(* IEC 61131-3 sources: ConveyorControl-with-PLC/4E_Gruppe1_Graf_Projekt1/Class/SafetyManager (part 3) *)

                    // change the command, because now we forward it to the receiver
                    pPara^.uiCmd := CMD_SM_SDO_TO_MODULE;

                    pHelpSafety^.pThis^.NewInst(pPara, #MyResult);
                    return;
                  else
                    pHelpSafety := pHelpSafety^.pNext;
                  end_if;
                end_while;
              end_if;
            end_if;

            pHelpPdo := pHelpPdo^.pNext;
          end_while;

          pHelpConfig := pHelpConfig^.pNext;
        end_while;
      end_if;
    end_if;

    // check if there is any interface frame domain optional and not available
    pHelpManaging := pFirstManagingInterfaceComponent;
    while pHelpManaging do
      if (pHelpManaging^.InfoBits.IsSynchron = 0) & (pHelpManaging^.InfoBits.IsOptional = 1) then
        // found one => no error here
        return;
      end_if;

      pHelpManaging := pHelpManaging^.pNext;
    end_while;

    // no optional interface domains missing => must be an error
    LogError("(SafetyManager::CheckTopSDO) Couldn't find InterfaceCRC. Check SafetyDesigner projects, maybe the interface variables do not match.");
    LogValue(pString:="SrcAddr: {0} / InterfaceCRC: {1}", Value:=pDO^.SrcAdr, Value2:=InterfaceCRC);
    ClassState := -8;

  // check if it's a local interface frame and we have no interface frame domains
  elsif (pCompDestPath^ = INTERFACE_CRC_MODE) then
    // after the mode byte we find the interface CRC
    InterfaceCRC := ((pCompDestPath + 1)$^HDINT)^;

    // search for the CRC
    pHelpSafety := NIL;
    if LocalIFNo then
      for i := 0 to (LocalIFNo-1) do
        if aLocalIFs[i].InterfaceCRC = InterfaceCRC then
          // found it
          pHelpSafety := aLocalIFs[i].pSafetyModule;
          exit;
        end_if;
      end_for;
    end_if;

    if pHelpSafety then
      // change the command, because now we forward it to the receiver
      pPara^.uiCmd := CMD_SM_SDO_TO_MODULE;

      pHelpSafety^.pThis^.NewInst(pPara, #MyResult);
    else
      // check the slave modules if there is one with the interface frame we need
      TargetSafetyNbr := 0;
      pHelpConfig := pConfigs;
      while pHelpConfig do
        pHelpSlave := pHelpConfig^.pFirstSlaveCfg;
        while pHelpSlave do

          if (pHelpSlave^.SlaveInfo.Info.IsInterface) & (pHelpSlave^.SlaveInfo.InterfaceCRC = InterfaceCRC) then
            // we have to add some additional information to the message

            (*
              Memory structure:
                1 Byte destination domain
                1 Byte IsInterfaceFrame (0/1)
                2 Byte length of uncompressed path
                x Byte uncompressed path
                x Byte SDO message
            *)

            MyPara.uiCmd := CMD_SM_TOP_SDO_TO_MODULE;
            MyPara.aPara[0] := sizeof(USINT) + sizeof(BOOL) + sizeof(UINT) + pHelpSlave^.SlaveInfo.PathLen + pPara^.aPara[0];

            if ud_SizeTempMemCy >= MyPara.aPara[0]$UDINT then
              pTempMem := pTempMemCy$^USINT;
            else
              LogError("(SafetyManager::CheckTopSDO) Temporary memory for cyclic task is too small!");
              LogValue(pString:="AvaliableMem: {0} / NeededMem: {1}", Value:=ud_SizeTempMemCy, Value2:=MyPara.aPara[0]$UDINT);
              return;
            end_if;

            TmpPathLen := pHelpSlave^.SlaveInfo.PathLen; // save some time with this local variable
            DomainChangeFound := FALSE;
            pHelp := pHelpSlave^.SlaveInfo.pPath + TmpPathLen - 2; // pointer on penultimate byte of path
            // search from the end for the last domain change
            for i := (TmpPathLen-2) to 3 by -1 do
              if pHelp^ = HWT_ESCAPE_DOMAIN then
                DomainChangeFound := TRUE;
                DestDomain := (pHelp + 1)^;
                exit;
              end_if;

              pHelp -= sizeof(USINT);
            end_for;

            // if there was no domainchange
            if DomainChangeFound = FALSE then
              // the master is the Dest
              DestDomain := (pHelpSlave^.SlaveInfo.pPath + 2)^;
            end_if;

            pHelp := pTempMem;

            // destination domain
            pHelp^ := DestDomain;
            pHelp += sizeof(USINT);

            // is it for an interface frame?
            pHelp^$BOOL := TRUE;
            pHelp += sizeof(BOOL);

            // length of uncompressed path
            pHelp^$UINT := TmpPathLen;
            pHelp += sizeof(UINT);

            // uncompressed path
            _memcpy(ptr1:=pHelp, ptr2:=pHelpSlave^.SlaveInfo.pPath, cntr:=TmpPathLen);
            pHelp += TmpPathLen;

            // SDO message
            _memcpy(ptr1:=pHelp, ptr2:=pDO, cntr:=pPara^.aPara[0]$UDINT);

            MyPara.aPara[1] := pTempMem$DINT;

            NewInst(#MyPara, #MyResult);

            // path can exist only once in a system
            return;
          end_if;

          pHelpSlave := pHelpSlave^.pNext;
        end_while;

        pHelpModule := pHelpConfig^.pFirstModuleCfg;
        while pHelpModule do
          if pHelpModule^.ModuleInfo.InterfaceCRC = InterfaceCRC then
            // if we found our target => forward the SDO to it
            TargetSafetyNbr := pHelpModule^.ModuleInfo.SafetyNbr;

            pHelpSafety := pFirstSafetyComponent;
            while pHelpSafety do
              // we compare the safety number
              if pHelpSafety^.SafetyNbr = TargetSafetyNbr then
                // change the command, because now we forward it to the receiver
                pPara^.uiCmd := CMD_SM_SDO_TO_MODULE;

                pHelpSafety^.pThis^.NewInst(pPara, #MyResult);

                return;
              end_if;

              pHelpSafety := pHelpSafety^.pNext;
            end_while;
          end_if;

          pHelpModule := pHelpModule^.pNext;
        end_while;

        pHelpConfig := pHelpConfig^.pNext;
      end_while;

      LogError("(SafetyManager::CheckTopSDO) Couldn't find target of SDO via TOP (Local Interface Frame)");
      LogValue(pString:="SrcAddr: {0} / InterfaceCRC: {1}", Value:=pDO^.SrcAdr, Value2:=InterfaceCRC);
    end_if;
  else
    // check if we have a module with this path
    pHelpConfig := pConfigs;
    while pHelpConfig do
      pHelpModule := pHelpConfig^.pFirstModuleCfg;
      while pHelpModule do
        if (To_StdLib.MemCmp(pCompDestPath, pHelpModule^.ModuleInfo.pCompPath, pHelpModule^.ModuleInfo.CompPathLen) = 0) then
          // we have to add some additional information to the message

          (*
            Memory structure:
              1 Byte destination domain
              1 Byte IsInterfaceFrame (0/1)
              2 Byte length of uncompressed path
              x Byte uncompressed path
              x Byte SDO message
          *)

          TmpPathLen := pHelpModule^.ModuleInfo.PathLen; // save some time with this local variable
          MyPara.uiCmd := CMD_SM_TOP_SDO_TO_MODULE;
          MyPara.aPara[0] := sizeof(USINT) + sizeof(BOOL) + sizeof(UINT) + TmpPathLen + pPara^.aPara[0];
          if ud_SizeTempMemCy >= MyPara.aPara[0]$UDINT then
            pTempMem := pTempMemCy$^USINT;
          else
            LogError("(SafetyManager::CheckTopSDO) Temporary memory for cyclic task is too small!");
            LogValue(pString:="AvaliableMem: {0} / NeededMem: {1}", Value:=ud_SizeTempMemCy, Value2:=MyPara.aPara[0]$UDINT);
            return;
          end_if;

          DomainChangeFound := FALSE;
          pHelp := pHelpModule^.ModuleInfo.pPath + TmpPathLen - 2; // pointer on penultimate byte of path
          // search from the end for the last domain change
          for i := (TmpPathLen-2) to 3 by -1 do
            if pHelp^ = HWT_ESCAPE_DOMAIN then
              DomainChangeFound := TRUE;
              DestDomain := (pHelp + 1)^;
              exit;
            end_if;

            pHelp -= sizeof(USINT);
          end_for;

          // if there was no domainchange
          if DomainChangeFound = FALSE then
            // the master is the Dest
            DestDomain := (pHelpModule^.ModuleInfo.pPath + 2)^;
          end_if;

          pHelp := pTempMem;

          // destination domain
          pHelp^ := DestDomain;
          pHelp += sizeof(USINT);

          // is it for an interface frame?
          pHelp^$BOOL := FALSE;
          pHelp += sizeof(BOOL);

          // length of uncompressed path
          pHelp^$UINT := TmpPathLen;
          pHelp += sizeof(UINT);

          // uncompressed path
          _memcpy(ptr1:=pHelp, ptr2:=pHelpModule^.ModuleInfo.pPath, cntr:=TmpPathLen);
          pHelp += TmpPathLen;

          // SDO message
          _memcpy(ptr1:=pHelp, ptr2:=pDO, cntr:=pPara^.aPara[0]$UDINT);

          MyPara.aPara[1] := pTempMem$DINT;

          NewInst(#MyPara, #MyResult);

          // path can exist only once in a system
          return;
        end_if;

        pHelpModule := pHelpModule^.pNext;
      end_while;

      if pHelpConfig^.SafetyNbr = pDO^.SrcAdr then
        pHelpSlave := pHelpConfig^.pFirstSlaveCfg;
        while pHelpSlave do
          if (To_StdLib.MemCmp(pCompDestPath, pHelpSlave^.SlaveInfo.pCompPath, pHelpSlave^.SlaveInfo.CompPathLen) = 0) then
            // we have to add some additional information to the message

            (*
              Memory structure:
                1 Byte destination domain
                1 Byte IsInterfaceFrame (0/1)
                2 Byte length of uncompressed path
                x Byte uncompressed path
                x Byte SDO message
            *)

            TmpPathLen := pHelpSlave^.SlaveInfo.PathLen; // save some time with this local variable
            MyPara.uiCmd := CMD_SM_TOP_SDO_TO_MODULE;
            MyPara.aPara[0] := sizeof(USINT) + sizeof(BOOL) + sizeof(UINT) + TmpPathLen + pPara^.aPara[0];
            if ud_SizeTempMemCy >= MyPara.aPara[0]$UDINT then
              pTempMem := pTempMemCy$^USINT;
            else
              LogError("(SafetyManager::CheckTopSDO) Temporary memory for cyclic task is too small!");
              LogValue(pString:="AvaliableMem: {0} / NeededMem: {1}", Value:=ud_SizeTempMemCy, Value2:=MyPara.aPara[0]$UDINT);
              return;
            end_if;

            DomainChangeFound := FALSE;
            pHelp := pHelpSlave^.SlaveInfo.pPath + TmpPathLen - 2; // pointer on penultimate byte of path
            // search from the end for the last domain change
            for i := (TmpPathLen-2) to 3 by -1 do
              if pHelp^ = HWT_ESCAPE_DOMAIN then
                DomainChangeFound := TRUE;
                DestDomain := (pHelp + 1)^;
                exit;
              end_if;

              pHelp -= sizeof(USINT);
            end_for;

            // if there was no domainchange
            if DomainChangeFound = FALSE then
              // the master is the Dest
              DestDomain := (pHelpSlave^.SlaveInfo.pPath + 2)^;
            end_if;

            pHelp := pTempMem;

            // destination domain
            pHelp^ := DestDomain;
            pHelp += sizeof(USINT);

            // is it for an interface frame?
            pHelp^$BOOL := FALSE;
            pHelp += sizeof(BOOL);

            // length of uncompressed path
            pHelp^$UINT := TmpPathLen;
            pHelp += sizeof(UINT);

            // uncompressed path
            _memcpy(ptr1:=pHelp, ptr2:=pHelpSlave^.SlaveInfo.pPath, cntr:=TmpPathLen);
            pHelp += TmpPathLen;

            // SDO message
            _memcpy(ptr1:=pHelp, ptr2:=pDO, cntr:=pPara^.aPara[0]$UDINT);

            MyPara.aPara[1] := pTempMem$DINT;

            NewInst(#MyPara, #MyResult);

            // path can exist only once in a system
            return;
          end_if;

          pHelpSlave := pHelpSlave^.pNext;
        end_while;
      end_if;

      pHelpConfig := pHelpConfig^.pNext;
    end_while;

    LogError("(SafetyManager::CheckTopSDO) Couldn't find destination of SDO. (Compressed Topology Path)");
    LogValue(pString:="SrcAddr: {0} / InterfaceCRC: {1}", Value:=pDO^.SrcAdr, Value2:=((pCompDestPath + 1)$^HDINT)^);

  end_if;

END_FUNCTION

FUNCTION SafetyManager::TopSDODest
	VAR_INPUT
		pPara 	: ^CmdStruct;
		pResult 	: ^results;
	END_VAR
	VAR_OUTPUT
		IsDestDomain 	: BOOL;
	END_VAR
  VAR
  	pHelpUSINT : ^USINT;
    PathLength : UINT;
    pPath : ^USINT;
    pHelpSafety : ^t_SafetyComponent;
  END_VAR

  IsDestDomain := FALSE;
(*
  Memory structure:
    1 Byte destination domain
    1 Byte IsInterfaceFrame (0/1)
    2 Byte length of uncompressed path
    x Byte uncompressed path
    x Byte SDO message
*)

  // check size (at least 1 byte for the destination domain + 2 byte for the path length + the header of the SDO message)
  if pPara^.aPara[0] > (sizeof(USINT) + sizeof(PathLength) + sizeof(SafetyCDIAS_Base::SDOHeader.StdHeader)) then
    pHelpUSINT := (pPara^.aPara[1])$^USINT;

    // domain
    pHelpUSINT += sizeof(USINT);

    // is it an interface frame info?
    pHelpUSINT += sizeof(BOOL);

    // path length
    PathLength := (pHelpUSINT$^UINT)^;
    pHelpUSINT += sizeof(UINT);

    // path
    pPath := pHelpUSINT;
    pHelpUSINT += PathLength;

    // pHelpUSINT points now to the SDO message

    // now we search the logged in modules for one with a matching topology path
    if pFirstSafetyComponent then

      pHelpSafety := pFirstSafetyComponent;
      while pHelpSafety do
        // we compare the last x byte (where x is the length of the local path including the domain)
        if pHelpSafety^.pPath & (To_StdLib.MemCmp(pHelpSafety^.pPath + 1, pPath + 2 + pPath^ - pHelpSafety^.pPath^, pHelpSafety^.pPath^) = 0) then
          pPara^.uiCmd := CMD_SM_SDO_TO_MODULE;
          pPara^.aPara[0] := pPara^.aPara[0] - (sizeof(USINT) + sizeof(PathLength) + PathLength);
          pPara^.aPara[1] := pHelpUSINT$DINT;

          pHelpSafety^.pThis^.NewInst(pPara, pResult);

          IsDestDomain := TRUE;
          return;
        end_if;

        pHelpSafety := pHelpSafety^.pNext;
      end_while;
    end_if;
  end_if;

END_FUNCTION

FUNCTION SafetyManager::PDOLengthCorrection
  VAR
  	pHelpConfig : ^t_CfgListElem;
    pHelpPDO    : ^t_PdoListElem;
    pHelpModule : ^t_ModuleListElem;
    pHelpSearchConfig : ^t_CfgListElem;
    FoundIt : BOOL;
    GotFirst : BOOL;
  END_VAR

  // with FSoE we use connections instead of the PDOs (PDOs are only remembered to check the optional state)
  if b_GotFSoEModules then
    return;
  end_if;

  GotFirst := FALSE;

  // check if there is a PDO with a zero length
  pHelpConfig := pConfigs;
  while pHelpConfig do
    pHelpPDO := pHelpConfig^.pFirstPdoCfg;
    while pHelpPDO do
      // remember the first PDO found as our act (to start from)
      if GotFirst = FALSE then
        GotFirst := TRUE;

        pActualSendCfg := pHelpConfig;
        pActualSendPDO := pHelpPDO;
      end_if;

      // if there is a PDO with no length
      if pHelpPDO^.PdoInfo.PdoLen = 0 then
        FoundIt := FALSE;
        pHelpSearchConfig := pConfigs;
        // search for the source module, because we use the length of it
        while pHelpSearchConfig & (FoundIt = FALSE) do
          pHelpModule := pHelpSearchConfig^.pFirstModuleCfg;
          while pHelpModule & (FoundIt = FALSE) do
            if pHelpModule^.ModuleInfo.PathLen = pHelpPDO^.PdoInfo.SourcePathLen then
              if (To_StdLib.MemCmp(pHelpModule^.ModuleInfo.pPath, pHelpPDO^.PdoInfo.pSourcePath, pHelpModule^.ModuleInfo.PathLen) = 0) then
                pHelpPDO^.PdoInfo.PdoLen := pHelpModule^.ModuleInfo.PdoOutLen;
                FoundIt := TRUE;
              end_if;
            end_if;

            pHelpModule := pHelpModule^.pNext;
          end_while;

          pHelpSearchConfig := pHelpSearchConfig^.pNext;
        end_while;
      end_if;

      pHelpPDO := pHelpPDO^.pNext;
    end_while;

    pHelpConfig := pHelpConfig^.pNext;
  end_while;

END_FUNCTION

FUNCTION SafetyManager::DoublePDOEntry
	VAR_INPUT
		NewPDO 	: t_PdoCfg;
		pNewCfg 	: ^t_CfgListElem;
	END_VAR
	VAR_OUTPUT
		IsDoubleEntry 	: BOOL;
	END_VAR
  VAR
  	pHelpCfg : ^t_CfgListElem;
    pHelpPdo : ^t_PdoListElem;
  END_VAR

  IsDoubleEntry := FALSE;

  // if it's our first config, there is no chance for a double PDO => check only if not first config
  if pNewCfg <> pConfigs then
    // otherwise: search all prior configs for the same PDO (source and destination path match)
    pHelpCfg := pConfigs;
    while pHelpCfg <> pNewCfg do
      pHelpPdo := pHelpCfg^.pFirstPdoCfg;
      while pHelpPdo do
        if (pHelpPdo^.PdoInfo.SourcePathLen = NewPDO.SourcePathLen) & (pHelpPdo^.PdoInfo.DestPathLen = NewPDO.DestPathLen) &
           (To_StdLib.MemCmp(pHelpPdo^.PdoInfo.pSourcePath, NewPDO.pSourcePath, NewPDO.SourcePathLen) = 0) &
           (To_StdLib.MemCmp(pHelpPdo^.PdoInfo.pDestPath, NewPDO.pDestPath, NewPDO.DestPathLen) = 0) then
          // we found the same PDO in a prior config
          IsDoubleEntry := TRUE;
          return;
        end_if;

        pHelpPdo := pHelpPdo^.pNext;
      end_while;

      pHelpCfg := pHelpCfg^.pNext;
    end_while;
  end_if;

END_FUNCTION

FUNCTION VIRTUAL SafetyManager::LogError
	VAR_INPUT
		e_msg 	: ^CHAR;
	END_VAR
  VAR
    sz_name : ARRAY [ 0..255 ] OF CHAR;
  END_VAR

  _GetObjName( this, #sz_name[ 0 ] );

  MyTrace(pFormat:="Object {0}: {1}", pTxt0:=(#sz_name[ 0 ])$^CHAR, pTxt1:= e_msg, pTxt2:=NIL);

END_FUNCTION

FUNCTION VIRTUAL SafetyManager::MyTrace
	VAR_INPUT
		pFormat 	: ^CHAR;
		pTxt0 	: ^CHAR;
		pTxt1 	: ^CHAR;
		pTxt2 	: ^CHAR;
	END_VAR
  VAR
    nLen      : UDINT;
    pChr      : ^CHAR;
    nTxt      : UDINT;
    nRpl      : UDINT;
    pTxt      : ^CHAR;
    pText     : ^CHAR;
    FormText  : ARRAY [0 .. 255] OF CHAR;
  END_VAR

  // this method is a workaround for the TRACE message limitation problem

  pText := #FormText[0];

  _memset(dest:=#FormText[0], usByte:=0, cntr:=256); // to keep the zero termination

  _strncpy(pText, pFormat, 250);
  nLen  := _strlen(pText);
  pChr  := pText;

  WHILE nLen DO
    IF pChr^ = '{' THEN         // works for the first 10 replacement texts (single digit numbers)
      nTxt  := (pChr+1)^ - '0';
      CASE nTxt OF
        0:  pTxt  := pTxt0;
        1:  pTxt  := pTxt1;
        2:  pTxt  := pTxt2;
      ELSE
        pTxt  := "INV";
      END_CASE;
      nRpl  := _strlen(pTxt);
      if nLen - 3 + nRpl > 250 then
        pTxt := "LEN";  // replace the replacement text with "LEN" to see that we're out of length for this string
        nRpl := 3;
      end_if;
      _memmove(pChr + nRpl, pChr + 3, nLen);
      _memcpy(pChr, pTxt, nRpl);
      pChr  += nRpl;  // next character to parse is after the replacement text
      nLen  -= 3;     // the remaining length of the format string is decremented by 3
      if nLen > 250 then  // catch overrun of nLen
        nLen := 0;
      end_if;
    ELSE
      pChr  += 1;
      nLen  -= 1;
    END_IF;
  END_WHILE;

  TRACE(#FormText[0]);
  if ( p_KernelLog ) then
    OS_KERNELLOG0(#FormText[0]);
  end_if;

END_FUNCTION

FUNCTION VIRTUAL SafetyManager::LogValue
	VAR_INPUT
		pString 	: ^CHAR;
		Value 	: UDINT;
		Value2 	: UDINT;
		Value3 	: UDINT;
	END_VAR
  VAR
    TempStr       : ARRAY [0..99] OF CHAR;
    TempStr2      : ARRAY [0..99] OF CHAR;
    TempStr3      : ARRAY [0..99] OF CHAR;
    TraceVal      : USINT;
    sz_name       : ARRAY [ 0..255 ] OF CHAR;
    TmpWithObjName: ARRAY [ 0..255 ] OF CHAR;
  END_VAR

  // number of values
  TraceVal := 1;

  _itoa(Value, #TempStr[0]);

  if pString <> NIL then
    _GetObjName( this, #sz_name[ 0 ] );
    _strcpy(dest:=#TmpWithObjName[0], src:="ObjectName ");
    _strcat(dest:=#TmpWithObjName[0], src:=#sz_name[0]);
    _strcat(dest:=#TmpWithObjName[0], src:=": ");
    _strcat(dest:=#TmpWithObjName[0], src:=pString);

    if Value2 <> 16#FFFFFFFF then
      _itoa(Value2, #TempStr2[0]);
      TraceVal += 1;
    end_if;

    if Value3 <> 16#FFFFFFFF then
      _itoa(Value3, #TempStr3[0]);
      TraceVal += 1;
    end_if;

    case TraceVal of
      1:MyTrace(pFormat:=#TmpWithObjName[0], pTxt0:=#TempStr[0], pTxt1:=NIL, pTxt2:=NIL);
      2:MyTrace(pFormat:=#TmpWithObjName[0], pTxt0:=#TempStr[0], pTxt1:=#TempStr2[0], pTxt2:=NIL);
      3:MyTrace(pFormat:=#TmpWithObjName[0], pTxt0:=#TempStr[0], pTxt1:=#TempStr2[0], pTxt2:=#TempStr3[0]);
    end_case;
  else
    MyTrace(pFormat:="<invalid string>", pTxt0:=NIL, pTxt1:=NIL, pTxt2:=NIL);
  end_if;

END_FUNCTION

FUNCTION SafetyManager::StoreInterfaceRoutingList
	VAR_INPUT
		pPara 	: ^CmdStruct;
		pResult 	: ^results;
		IsFSoE 	: BOOL;
	END_VAR
  VAR
  	pHelpManaging : ^t_ManagingComponent;
    EntryNo       : USINT;
    i             : UDINT;
    pHelp         : ^t_InterfaceFrameInfo;
    ActOffset     : UDINT;
    pHelpFSoE     : ^t_IFConnectionInfo;
    j             : UDINT;
    GenerateNo    : USINT;
    OldFSoENo     : DINT;
  END_VAR

  if IsFSoE then

    // if we already have different data from this management component => delete the old stuff first
    if IFFSoENo then
      OldFSoENo := IFFSoENo$DINT;

      // remove the existing stuff of this managing component
      for i$DINT := (OldFSoENo-1) to 0 by -1 do
        // check if it's from the same managing component
        if aIFFSoEInfos[i].pManaging^.pThis$DINT = pPara^.aPara[2] then
          // remove it

          // move the following blocks over this one (if it's not the last)
          if i$UDINT < IFFSoENo-1 then
            for j := i to (IFFSoENo-2) do
              aIFFSoEInfos[j] := aIFFSoEInfos[j+1];
            end_for;
          end_if;
          IFFSoENo -= 1;
        end_if;
      end_for;
    end_if;

    EntryNo := ((pPara^.aPara[0] - sizeof(t_IFInfoFSoE.IsResponse)) / sizeof(t_IFConnectionInfo))$USINT;
    if (EntryNo + IFFSoENo <= MAX_MODULES_IN_OTHER_DOMAINS) then
      ActOffset := 0;
      pHelpManaging := pFirstManagingInterfaceComponent;
      while pHelpManaging do
        // if we found the sender of this list in our list of interfaceframe components, remember the safety numbers
        if pHelpManaging^.pThis$DINT = pPara^.aPara[2] then
          if EntryNo then

            // set the help pointer to the first entry of the interface frame info array
            pHelpFSoE := pPara^.aPara[1]$^t_IFConnectionInfo + sizeof(BOOL);
            for i := 0 to (EntryNo-1) do
              pHelpManaging^.ModuleInfo[i].SafetyNbr := pHelpFSoE^.SafetyNbr;

              if pHelpFSoE^.Flags.IsMaster then
                pHelpManaging^.ModuleInfo[i].InfoBits.IsFSoEMaster := TRUE;
                pHelpManaging^.ModuleInfo[i].InfoBits.IsFSoESlave  := FALSE;
              else
                pHelpManaging^.ModuleInfo[i].InfoBits.IsFSoEMaster := FALSE;
                pHelpManaging^.ModuleInfo[i].InfoBits.IsFSoESlave  := TRUE;
              end_if;

              // we save the whole info for PDO/SDO routing
              aIFFSoEInfos[IFFSoENo].FromOtherSide := pHelpFSoE^;
              aIFFSoEInfos[IFFSoENo].FromOtherSide.FollowUps := 0; // only relevant for the transfer to this domain
              aIFFSoEInfos[IFFSoENo].pManaging := pHelpManaging;

              IFFSoENo += 1;

              if pHelpFSoE^.FollowUps then
                GenerateNo := pHelpFSoE^.FollowUps;
                for j := 1 to GenerateNo do
                  // we save the whole info for PDO/SDO routing
                  aIFFSoEInfos[IFFSoENo].FromOtherSide := pHelpFSoE^;
                  aIFFSoEInfos[IFFSoENo].FromOtherSide.FollowUps := 0; // only relevant for the transfer to this domain
                  aIFFSoEInfos[IFFSoENo].pManaging := pHelpManaging;

                  IFFSoENo += 1;
                end_for;
              end_if;

              pHelpFSoE += sizeof(t_IFConnectionInfo);
            end_for;
          end_if;

          pHelpManaging^.ModuleNo := EntryNo;

          pHelpManaging^.InfoBits.GotIFInfo := TRUE;
          return;
        end_if;

        pHelpManaging := pHelpManaging^.pNext;
      end_while;
    else
      LogError("(SafetyManager::StoreInterfaceRoutingList) Invalid size of configuration (FSoE)");
    end_if;
  else
    EntryNo := ((pPara^.aPara[0] - sizeof(t_IFInfo.IsResponse)) / sizeof(t_InterfaceFrameInfo))$USINT;

    if (EntryNo + InterfaceFrameNo <= MAX_MODULES_IN_OTHER_DOMAINS) then
      ActOffset := 0;
      pHelpManaging := pFirstManagingInterfaceComponent;
      while pHelpManaging do
        // if we found the sender of this list in our list of interfaceframe components, remember the safety numbers
        if pHelpManaging^.pThis$DINT = pPara^.aPara[2] then
          if EntryNo then
            // set the help pointer to the first entry of the interface frame info array
            pHelp := pPara^.aPara[1]$^t_InterfaceFrameInfo + sizeof(BOOL);
            for i := 0 to (EntryNo-1) do
              // we save the module info's with the domain interface module for TDO/SDO routing
              pHelpManaging^.ModuleInfo[i] := pHelp^.ModuleInfo;

              // we also save the whole info for PDO routing
              aInterfaceFrameInfos[InterfaceFrameNo] := pHelp^;

              // only for IFs where the communication partner is the source
              if aInterfaceFrameInfos[InterfaceFrameNo].IFPdoLen then
                aInterfaceFrameInfos[InterfaceFrameNo].OffsetInDomainModule := ActOffset;
                ActOffset += aInterfaceFrameInfos[InterfaceFrameNo].IFPdoLen;
              end_if;

              InterfaceFrameNo += 1;

              pHelp += sizeof(t_InterfaceFrameInfo);
            end_for;
          end_if;

          pHelpManaging^.ModuleNo := EntryNo;

          pHelpManaging^.InfoBits.GotIFInfo := TRUE;
          return;
        end_if;

        pHelpManaging := pHelpManaging^.pNext;
      end_while;
    else
      LogError("(SafetyManager::StoreInterfaceRoutingList) Invalid size of configuration");
    end_if;
  end_if;

END_FUNCTION

FUNCTION SafetyManager::AllInterfaceCfgsArrived
	VAR_OUTPUT
		AllReady 	: BOOL;
	END_VAR
  VAR
    pHelpManaging : ^t_ManagingComponent;
  END_VAR

  AllReady := TRUE;

  // check if we have the safety numbers for every interface managing module in the system
  pHelpManaging := pFirstManagingInterfaceComponent;
  while pHelpManaging do
    if pHelpManaging^.InfoBits.IsSynchron & (pHelpManaging^.InfoBits.GotIFInfo = FALSE) then
      AllReady := FALSE;
      return;
    end_if;

    pHelpManaging := pHelpManaging^.pNext;
  end_while;

END_FUNCTION

FUNCTION SafetyManager::SendInterfaceConfigs
	VAR_INPUT
		DestinationThis 	: pVirtualBase;(* := NIL *)
		IsResponse 	: BOOL;(* := FALSE *)
		IsFSoE 	: BOOL;
	END_VAR
  VAR
    pHelpCfg                  : ^t_CfgListElem;
    pHelpModule               : ^t_ModuleListElem;
    pHelpPdo                  : ^t_PdoListElem;
    pHelpConnection           : ^t_FSoEConnectionDetails;
    MyPara                    : CmdStruct;
    MyResult                  : results;
    TmpIFInfo                 : t_IFInfo;
    ModuleInfoNo              : USINT;
    i                         : UDINT;
    pActCRC                   : ^HDINT;
    TmpIFConn                 : t_IFInfoFSoESend;
    pLastReferenceConnection  : ^t_IFConnectionInfo;
  END_VAR

  // collect the safety numbers of this system
  ModuleInfoNo := 0;

  if IsFSoE then
    //reset memory => now 0 is an invalid safety number (= unused element of the array)
    _memset(dest:=#TmpIFConn, usByte:=0, cntr:=sizeof(t_IFInfoFSoESend));
    TmpIFConn.IsResponse := IsResponse;

    pLastReferenceConnection  := NIL;

    // if not all configs available, create and send the available data
    if (LocalCPUCfgNo <> LocalCPUNo) then
      // check FSoE Connections in the available configs
      pHelpCfg := pConfigs;
      while pHelpCfg do
        pHelpConnection := pHelpCfg^.pFirstFSoEConnection;
        while pHelpConnection do
          // only interface connections are relevant
          if pHelpConnection^.Flags.IsInterfaceConnection then
            if pLastReferenceConnection & (pHelpConnection^.SlaveAddress = pLastReferenceConnection^.SlaveAddress) &
               (pHelpConnection^.Flags.IsMaster = pLastReferenceConnection^.Flags.IsMaster) then
              pLastReferenceConnection^.FollowUps += 1;
            else
              // add the modules to the info message
              TmpIFConn.aConnectionInfos[ModuleInfoNo].Flags            := pHelpConnection^.Flags;
              TmpIFConn.aConnectionInfos[ModuleInfoNo].SlaveAddress     := pHelpConnection^.SlaveAddress;
              TmpIFConn.aConnectionInfos[ModuleInfoNo].SafetyNbr        := pHelpConnection^.OwnerSafetyNbr;
              TmpIFConn.aConnectionInfos[ModuleInfoNo].MasterReadSize   := pHelpConnection^.MasterReadSize;
              TmpIFConn.aConnectionInfos[ModuleInfoNo].MasterWriteSize  := pHelpConnection^.MasterWriteSize;
              TmpIFConn.aConnectionInfos[ModuleInfoNo].FollowUps        := 0;

              // some data are only available at the master
              if pHelpConnection^.Flags.IsMaster then
                // no follow ups for master connections
                pLastReferenceConnection                                := NIL;

                TmpIFConn.aConnectionInfos[ModuleInfoNo].ConnectionID   := pHelpConnection^.ConnectionID;
              else
                // update this value for the next connections with the same settings to save a lot of memory
                pLastReferenceConnection                                := #TmpIFConn.aConnectionInfos[ModuleInfoNo];

                TmpIFConn.aConnectionInfos[ModuleInfoNo].ConnectionID   := 0;
              end_if;

              if pHelpConnection^.SlavePathCompLen & pHelpConnection^.pSlavePathComp then
                TmpIFConn.aConnectionInfos[ModuleInfoNo].InterfaceCRC := (pHelpConnection^.pSlavePathComp$^HDINT + 1)^;
              else
                TmpIFConn.aConnectionInfos[ModuleInfoNo].InterfaceCRC := 0;
              end_if;

              ModuleInfoNo += 1;
            end_if;
          end_if;

          pHelpConnection := pHelpConnection^.pNext;
        end_while;

        pHelpCfg := pHelpCfg^.pNext;
      end_while;
    else
      // check FSoE Connections in the sorted list
      pHelpConnection := pSortedConnections;
      while pHelpConnection do
        // only interface connections are relevant
        if pHelpConnection^.Flags.IsInterfaceConnection then
          if pLastReferenceConnection & (pHelpConnection^.SlaveAddress = pLastReferenceConnection^.SlaveAddress) &
             (pHelpConnection^.Flags.IsMaster = pLastReferenceConnection^.Flags.IsMaster) then
            pLastReferenceConnection^.FollowUps += 1;
          else
            // add the modules to the info message
            TmpIFConn.aConnectionInfos[ModuleInfoNo].Flags            := pHelpConnection^.Flags;
            TmpIFConn.aConnectionInfos[ModuleInfoNo].SlaveAddress     := pHelpConnection^.SlaveAddress;
            TmpIFConn.aConnectionInfos[ModuleInfoNo].SafetyNbr        := pHelpConnection^.OwnerSafetyNbr;
            TmpIFConn.aConnectionInfos[ModuleInfoNo].MasterReadSize   := pHelpConnection^.MasterReadSize;
            TmpIFConn.aConnectionInfos[ModuleInfoNo].MasterWriteSize  := pHelpConnection^.MasterWriteSize;
            TmpIFConn.aConnectionInfos[ModuleInfoNo].FollowUps        := 0;

            // some data are only available at the master
            if pHelpConnection^.Flags.IsMaster then
              // no follow ups for master connections
              pLastReferenceConnection                                := NIL;

              TmpIFConn.aConnectionInfos[ModuleInfoNo].ConnectionID   := pHelpConnection^.ConnectionID;
            else
              // update this value for the next connections with the same settings to save a lot of memory
              pLastReferenceConnection                                := #TmpIFConn.aConnectionInfos[ModuleInfoNo];

              TmpIFConn.aConnectionInfos[ModuleInfoNo].ConnectionID   := 0;
            end_if;

            if pHelpConnection^.SlavePathCompLen & pHelpConnection^.pSlavePathComp then
              TmpIFConn.aConnectionInfos[ModuleInfoNo].InterfaceCRC := (pHelpConnection^.pSlavePathComp$^HDINT + 1)^;
            else
              TmpIFConn.aConnectionInfos[ModuleInfoNo].InterfaceCRC := 0;
            end_if;

            ModuleInfoNo += 1;
          end_if;
        end_if;

        pHelpConnection := pHelpConnection^.pNextSorted;
      end_while;
    end_if;

    CheckLocalSlaveAddresses();

    if b_AllLocalSlaveAddressesValid then
      MyPara.uiCmd := CMD_SM_IF_MODULE_INFO_FSOE_OK;
    else
      MyPara.uiCmd := CMD_SM_IF_MODULE_INFO_FSOE;
    end_if;

    MyPara.aPara[0] := ModuleInfoNo * sizeof(t_IFConnectionInfo) + sizeof(t_IFInfoFSoE.IsResponse);
    MyPara.aPara[1] := (#TmpIFConn)$DINT;
  else
    // browse through the configs
    TmpIFInfo.IsResponse := IsResponse;

    pHelpCfg := pConfigs;
    while pHelpCfg do
      pHelpPdo := pHelpCfg^.pFirstPdoCfg;
      while pHelpPdo do
        // if it's a interface broadcast
        if pHelpPdo^.PdoInfo.Info.IFBroadCast then
          // search for the source module
          pHelpModule := pHelpCfg^.pFirstModuleCfg;
          while pHelpModule do
            // if it's an interface source and the interface CRC matches the one of our PDO => Bingo! But to be sure we check also the path length and the path itself
            if pHelpModule^.ModuleInfo.Info.IsInterfaceSource & (pHelpModule^.ModuleInfo.InterfaceCRC = pHelpPdo^.PdoInfo.InterfaceCRC) &
              (pHelpModule^.ModuleInfo.PathLen = pHelpPdo^.PdoInfo.SourcePathLen) &
              (To_StdLib.MemCmp(pHelpModule^.ModuleInfo.pPath, pHelpPdo^.PdoInfo.pSourcePath, pHelpPdo^.PdoInfo.SourcePathLen) = 0) then

              TmpIFInfo.aModuleInfos[ModuleInfoNo].InterfaceCRC          := pHelpModule^.ModuleInfo.InterfaceCRC;
              TmpIFInfo.aModuleInfos[ModuleInfoNo].IFPdoLen              := pHelpPdo^.PdoInfo.PdoLen;
              TmpIFInfo.aModuleInfos[ModuleInfoNo].OffsetInDomainModule  := 0; // the correct offset is calculated in the receiver
              TmpIFInfo.aModuleInfos[ModuleInfoNo].ModuleInfo.SafetyNbr  := pHelpModule^.ModuleInfo.SafetyNbr;

              ModuleInfoNo += 1;
            end_if;

            pHelpModule := pHelpModule^.pNext;
          end_while;
        end_if;

        pHelpPdo := pHelpPdo^.pNext;
      end_while;

      // check the modules of the actual config if there are interface frame destinations (needed for unidirectional communication, otherwise the SDO routing would fail)
      pHelpModule := pHelpCfg^.pFirstModuleCfg;
      while pHelpModule do
        // if it's a interface destination
        if pHelpModule^.ModuleInfo.Info.IsInterfaceDest then
          pActCRC := pHelpModule^.ModuleInfo.pDestCRCs;
          for i := 0 to (pHelpModule^.ModuleInfo.DestCRCNo-1) do
            TmpIFInfo.aModuleInfos[ModuleInfoNo].InterfaceCRC          := pActCRC^;
            TmpIFInfo.aModuleInfos[ModuleInfoNo].IFPdoLen              := 0; // we don't know the length here, we're only the receiver
            TmpIFInfo.aModuleInfos[ModuleInfoNo].OffsetInDomainModule  := 0; // the correct offset is calculated in the receiver
            TmpIFInfo.aModuleInfos[ModuleInfoNo].ModuleInfo.SafetyNbr  := pHelpModule^.ModuleInfo.SafetyNbr;
            TmpIFInfo.aModuleInfos[ModuleInfoNo].ModuleInfo.InfoBits$UDINT := 0;

            pActCRC += sizeof(HDINT);
            ModuleInfoNo += 1;
          end_for;
        end_if;

        pHelpModule := pHelpModule^.pNext;
      end_while;

      pHelpCfg := pHelpCfg^.pNext;
    end_while;

    MyPara.uiCmd := CMD_SM_IF_MODULE_INFO;
    MyPara.aPara[0] := ModuleInfoNo * sizeof(t_InterfaceFrameInfo) + sizeof(TmpIFInfo.IsResponse);
    MyPara.aPara[1] := (#TmpIFInfo)$DINT;
  end_if;

  // if we have only 1 destination => sent it to this destination
  if DestinationThis then
    DestinationThis^.NewInst(#MyPara, #MyResult);
  else
    // otherwise send our safety numbers to every interface managing module in the system
    TellAllInterfaceManagingModules(#MyPara, #MyResult);
  end_if;

END_FUNCTION

FUNCTION SafetyManager::GetIFInfoByCRC
	VAR_INPUT
		InterfaceCRC 	: HDINT;
		pMemOffset 	: ^UDINT;
		pLength 	: ^USINT;
	END_VAR
	VAR_OUTPUT
		SafetyNbr 	: HDINT;
	END_VAR
  VAR
    i : UDINT;
  END_VAR

  SafetyNbr := 0;

  if InterfaceFrameNo then
    for i := 0 to (InterfaceFrameNo-1) do
      // if we found the interface CRC and it's a interface frame we receive (the sender adds the length)
      if (aInterfaceFrameInfos[i].InterfaceCRC = InterfaceCRC) & aInterfaceFrameInfos[i].IFPdoLen then
        SafetyNbr := aInterfaceFrameInfos[i].ModuleInfo.SafetyNbr;
        // check if pointers are valid
        if pMemOffset & pLength then
          pMemOffset^ := aInterfaceFrameInfos[i].OffsetInDomainModule;
          pLength^    := aInterfaceFrameInfos[i].IFPdoLen;
        end_if;
        return;
      end_if;
    end_for;

    if SafetyNbr = 0 then
      LogError("(SafetyManager::GetIFInfoByCRC) Safetynumber of Interface-Frame source couldn't be found in the list");
    end_if;
  end_if;

END_FUNCTION

FUNCTION SafetyManager::SetTimeout

  ud_InitTimeOut := ops.tAbsolute;

END_FUNCTION

FUNCTION SafetyManager::CheckTimeout

  // if the step took too long
  if (OPS.tAbsolute - ud_InitTimeOut) > T_INIT_TIMEOUT then
    // show the possible error in the log/trace and restart the time for timeout
    case InitSSW of
//**********************************************************************************************************************************************************
      _FirstWait4SynchronSubdomains:
        LogError("Timeout in Initialisation of SafetyManager while waiting first time for subdomains to get synchron!");
//**********************************************************************************************************************************************************
      _Wait4FSoEConnectionsLocal:
        LogError("Timeout in Initialisation of SafetyManager while waiting for the local FSoE connections to get initialized!");
//**********************************************************************************************************************************************************
      _Wait4SynchronSubdomains:
        LogError("Timeout in Initialisation of SafetyManager while waiting for subdomains to get synchron!");
//**********************************************************************************************************************************************************
      _Wait4ConfigFlush:
        LogError("Timeout in Initialisation of SafetyManager while waiting for the slave domains to send their safety numbers of safety cpus and if they can handle the new time sync method!");
//**********************************************************************************************************************************************************
      _Wait4CPUConfigs:
        LogError("Timeout in Initialisation of SafetyManager while waiting for all available cpu configurations!");
//**********************************************************************************************************************************************************
      _Wait4InterfaceConfigs:
        LogError("Timeout in Initialisation of SafetyManager while waiting for module informations from another domain needed for interface frame communication!");
//**********************************************************************************************************************************************************
      _Wait4FSoEConnectionsExternal:
        LogError("Timeout in Initialisation of SafetyManager while waiting for the external FSoE connections to get initialized!");
//**********************************************************************************************************************************************************
      _Wait4UnsafeConfigAck:
        LogError("Timeout in Initialisation of SafetyManager while waiting for an unsafe variable configuration acknowledgment of another domain!");
//**********************************************************************************************************************************************************
      _Wait4PDOAcks:
        LogError("Timeout in Initialisation of SafetyManager while waiting for a pdo configuration acknowledgment!");
//**********************************************************************************************************************************************************
    end_case;

    // this error gets quitted if initialisation finishes
    ClassState := -11;

    ud_InitTimeOut := ops.tAbsolute;
  end_if;

END_FUNCTION

FUNCTION SafetyManager::AllNonOptionalIFDomainsSynchron
	VAR_OUTPUT
		EverythingSynchron 	: BOOL;
	END_VAR
  VAR
  	pHelpManaging : ^t_ManagingComponent;
    pHelpConfig : ^t_CfgListElem;
    pHelpPdo : ^t_PdoListElem;
    TempCfg : t_PdoCfg;
		MyPara 	  : CmdStruct;
		MyResult	: results;
  END_VAR

  EverythingSynchron := TRUE;

  MyPara.uiCmd := CMD_SM_SYNC_CHECK;

  // check for all interface frame PDOs in the configurations if the corresponding domain managing module is synchron
  pHelpConfig := pConfigs;
  while pHelpConfig do
    pHelpPdo := pHelpConfig^.pFirstPdoCfg;
    while pHelpPdo do
      TempCfg := pHelpPdo^.PdoInfo;
      // if it's an interface  PDO, no double entry and not optional => it has to be synchron!
      if (TempCfg.Info.IsInterfacePDO = TRUE) & (TempCfg.Info.DoublePDOEntry = FALSE) & (TempCfg.Info.IsOptional = FALSE) then
        pHelpManaging := pFirstManagingInterfaceComponent;
        while pHelpManaging do
          // we found the corresponding domain managing module
          if (pHelpManaging^.InfoBits.IsOptional = FALSE) &
            ((To_StdLib.MemCmp(pHelpManaging^.pModulePath, TempCfg.pSourcePath, TempCfg.SourcePathLen) = 0) |
             (To_StdLib.MemCmp(pHelpManaging^.pModulePath, TempCfg.pDestPath, TempCfg.DestPathLen) = 0)) then

            // if any of those is not synchron, stop searching
            if pHelpManaging^.pThis^.NewInst(#MyPara, #MyResult) = ERROR then
              EverythingSynchron := FALSE;
              return;
            end_if;

            exit;
          end_if;

          pHelpManaging := pHelpManaging^.pNext;
        end_while;
      end_if;

      pHelpPdo := pHelpPdo^.pNext;
    end_while;

    pHelpConfig := pHelpConfig^.pNext;
  end_while;

END_FUNCTION

FUNCTION VIRTUAL SafetyManager::GetThisViaServerName
	VAR_INPUT
		pObjectDotServer 	: ^CHAR;
	END_VAR
	VAR_OUTPUT
		ThisPtr 	: pVoid;
	END_VAR
  VAR
    ChannelMode : CHMODE;
  END_VAR

  ThisPtr := NIL;

  if pObjectDotServer = NIL then
    return;
  end_if;

  // get thispointer to server via name
  ChannelMode := _LookUpEmbed_C(pObjectDotServer, #ThisPtr, NIL);

  // check if it's a server
  case ChannelMode of
    _CH_CMD,
    _CH_SVR:

  else
    ThisPtr := NIL;
    LogError(e_msg:="(SafetyManager::GetThisViaServerName) Couldn't get thispointer of server:");
    LogError(e_msg:=pObjectDotServer);
  end_case;

END_FUNCTION

FUNCTION SafetyManager::GetNewMovDO
	VAR_OUTPUT
		Index 	: INT;
	END_VAR
//  VAR
//  	sd_retval : DINT;
//  END_VAR

  Index := -1;

  if CopyCmdsUsed < MAX_PDO_COPY_CMDS then
    // check if there is one available but not used
    if CopyCmdsUsed < CopyCmdsAvailable then
      Index := CopyCmdsUsed;
      CopyCmdsUsed += 1;
    else
      // we have to create a new one

(*
// connection to varan manager required
      // add data object to copy our data
      sd_retval := pVaranManager^.AddMovDO(ud_dol_type:=VARAN_DOL_ISO
                                         , p_ud_handle:=(#aCopyCmds[CopyCmdsAvailable].pHandle)$^UDINT
                                         , p_ud_MovSettings:=( #aCopyCmds[CopyCmdsAvailable].pSettings)$^UDINT
                                         , ud_type := VM_PRIORITY_2
                                         );

      //look for an error
      if ( sd_retval <> 0 ) then
        ClassState := -9;
        LogError("(SafetyManager::GetNewMovDO) Failed to add a new copy command to the VaranManager!");
        return;
      end_if;
*)
      aCopyCmds[CopyCmdsAvailable].b_Ready4Action := FALSE;

      Index := CopyCmdsAvailable;

      CopyCmdsAvailable += 1;
      CopyCmdsUsed += 1;
    end_if;
  else
    LogError("Maximum of possible PDO copy commands reached!");
  end_if;

END_FUNCTION

FUNCTION SafetyManager::CheckCPUConfigs
	VAR_OUTPUT
		ConfigsOK 	: BOOL;
	END_VAR
  VAR
  	pHelpManaging   : ^t_ManagingComponent;
    pSourceManaging : ^t_ManagingComponent;
    pHelpConfig     : ^t_CfgListElem;
    pHelpPdo        : ^t_PdoListElem;
    pLastPdo        : ^t_PdoListElem;
    IsSource        : DINT;
    PDOCount : UDINT;
  END_VAR

  // before we go into the usual check routine, we have to ensure that we have enough virtual PDOs for writing interface frames (config holds a broadcast and we have to look for possible target modules)
  CreateVirtualPDOs();

  // initialize with true (normal case is that everything is ok => now we check for errors)
  ConfigsOK := TRUE;

  PDOCount := 0;

  // check if all non-optional modules are available and all corresponding domain managing module are synchron (if necessary)
  pHelpConfig := pConfigs;
  while pHelpConfig do
    pLastPdo := NIL;
    pHelpPdo := pHelpConfig^.pFirstPdoCfg;
    while pHelpPdo do
      // if it's an interface frame and no broadcast frame
      if pHelpPdo^.PdoInfo.Info.IsInterfacePDO then
        if (pHelpPdo^.PdoInfo.Info.IFBroadCast = FALSE) then

          // check if we have already added the domain interface to the IF List
          IsSource := -1; // -1 = not found, 0 = destination, 1 = source
          pSourceManaging := NIL;
          pHelpManaging := pFirstManagingInterfaceComponent;
          while pHelpManaging do
            // if source or destination of the PDO matches our managing module path => it's an interface frame to/from this domain
            if (To_StdLib.MemCmp(pHelpManaging^.pModulePath, pHelpPdo^.PdoInfo.pSourcePath, pHelpPdo^.PdoInfo.SourcePathLen) = 0) then
              pSourceManaging := pHelpManaging;
              IsSource := 1;
              exit;
            elsif (To_StdLib.MemCmp(pHelpManaging^.pModulePath, pHelpPdo^.PdoInfo.pDestPath, pHelpPdo^.PdoInfo.DestPathLen) = 0) then
              IsSource := 0;
              exit;
            end_if;

            pHelpManaging := pHelpManaging^.pNext;
          end_while;

          // if we got a source managing module and it isn't synchron
          if pSourceManaging then
            // if this pdo is not optional => the source module also isn't
            if pHelpPdo^.PdoInfo.Info.IsOptional = FALSE then
              pSourceManaging^.InfoBits.IsOptional := FALSE;
            end_if;

            if (pSourceManaging^.InfoBits.IsSynchron = FALSE) then
              if pHelpPdo^.PdoInfo.Info.IsOptional then
                // ignore it
  //              LogError("Info: Optional interface frame can't be received, because source domain is not connected or not synchron");

                // remove the PDO from the list (if not the receiver module would wait endless for the PDO and we can't send the set bus ready to quit errors of local PDOs)
                if pLastPdo then
                  // if we had already a PDO before in this configuration we have to skip the removed PDO with the next pointer
                  pLastPdo^.pNext := pHelpPdo^.pNext;

                  To_StdLib.Free(pHelpPdo^.PdoInfo.pSourcePath);
                  To_StdLib.Free(pHelpPdo^.PdoInfo.pDestPath);
                  To_StdLib.Free(pHelpPdo);

                  pHelpPdo := pLastPdo;
                else
                  // if it was the first PDO, we have to correct the first pointer
                  pHelpConfig^.pFirstPdoCfg := pHelpPdo^.pNext;

                  To_StdLib.Free(pHelpPdo^.PdoInfo.pSourcePath);
                  To_StdLib.Free(pHelpPdo^.PdoInfo.pDestPath);
                  To_StdLib.Free(pHelpPdo);

                  pHelpPdo := pHelpConfig^.pFirstPdoCfg;
                end_if;

                if pHelpPdo = NIL then
                  exit;
                end_if;
              else
                // non-optional interface frame domain missing => error
                LogError("ERROR! Non-Optional interface frame can't be received, because domain is not connected");
                ConfigsOK := FALSE;
                ClassState := -10;
              end_if;
            end_if;
          end_if;
        end_if;
      end_if;

      PDOCount += 1;

      pLastPdo := pHelpPdo;
      pHelpPdo := pHelpPdo^.pNext;
    end_while;

    pHelpConfig := pHelpConfig^.pNext;
  end_while;

  // if now PDOs found => reset the act ID to show that there are none
  if PDOCount = 0 then
    ActPDO_ID := 0;
  end_if;

END_FUNCTION

FUNCTION SafetyManager::RemoveLocalCPUCfg
	VAR_INPUT
		SafetyNumber 	: HDINT;
	END_VAR
  VAR
  	pHelpCfg    : ^t_LocalCfgListElem;
    i : UDINT;
  END_VAR

  if LocalCPUCfgNo then
    pHelpCfg := pFirstLocalCPUCfg;
    for i := 0 to (LocalCPUCfgNo-1) do
      if pHelpCfg^.SafetyNbr = SafetyNumber then
        // found it => deactivate it
        pHelpCfg^.ConfigSize := 0;
        pHelpCfg^.ConfigSent2Master := FALSE;
        exit;
      end_if;

      pHelpCfg := pHelpCfg^.pNext;
    end_for;
  end_if;

END_FUNCTION

FUNCTION SafetyManager::ClearRoutingInformations
  VAR
  	MyPara : CmdStruct;
    MyResult : results;
    pHelpManaging : ^t_ManagingComponent;
    i : UDINT;
    pHelpCfg      : ^t_LocalCfgListElem;
  END_VAR

  // we're flushin our stuff here

  // reset number of memorized safe cpu numbers
  SafeCPU_Nbr_No := 0;

  // set ID to zero for the next mapping assignment
  ActPDO_ID := 0;

  // reset interface frameno
  InterfaceFrameNo := IFFSoENo := 0;

  // reset local interface frameno
  LocalIFNo := 0;

  // clear configurations of safety-cpus
  FreeCfgLists();

  // clear number of copy DOs used
  CopyCmdsUsed := 0;

  // reset memory usage for isochronous transfer (the values are set when distributing the PDOs)
  MyPara.aPara[0] := 0;
  pHelpManaging := pFirstManagingInterfaceComponent;
  while pHelpManaging do
    pHelpManaging^.PDOReadMemUsed := 0;
    pHelpManaging^.PDOWriteMemUsed := 0;

    MyPara.uiCmd := CMD_SM_PDO_MEM_USAGE_WR;
    pHelpManaging^.pThis^.NewInst(#MyPara, #MyResult);

    MyPara.uiCmd := CMD_SM_PDO_MEM_USAGE_RD;
    pHelpManaging^.pThis^.NewInst(#MyPara, #MyResult);

    pHelpManaging^.InfoBits.HasBeenFlushed      := FALSE;
    pHelpManaging^.InfoBits.NewTimeSyncPossible := FALSE;
    pHelpManaging^.InfoBits.SubDomainsSynchron  := FALSE;
    pHelpManaging^.InfoBits.GotIFInfo           := FALSE;
    pHelpManaging^.InfoBits.LocalConfigReady    := FALSE;
    pHelpManaging^.InfoBits.IsOptional          := TRUE;  // initialize with true, later in the init process (CheckCPUConfigs) it's checked and corrected if necessary
    // synchron bit is already true at this time (or the timeout has expired)

    pHelpManaging^.DomainNr := 16#FF;

    pHelpManaging^.SubDomainsUsed := 0;
    _memset(dest:=#pHelpManaging^.SubDomainNr, usByte:=16#FF, cntr:=sizeof(pHelpManaging^.SubDomainNr));

    pHelpManaging^.ModuleNo := 0;
    _memset(dest:=#pHelpManaging^.ModuleInfo, usByte:=16#00, cntr:=sizeof(pHelpManaging^.ModuleInfo));

    pHelpManaging := pHelpManaging^.pNext;
  end_while;

  // all local cpu configs have to be sent again on reconnect
  if LocalCPUCfgNo then
    pHelpCfg := pFirstLocalCPUCfg;
    for i := 0 to (LocalCPUCfgNo-1) do
      pHelpCfg^.ConfigSent2Master := FALSE;

      pHelpCfg := pHelpCfg^.pNext;
    end_for;
  end_if;

END_FUNCTION

FUNCTION SafetyManager::CheckPDORecycle
	VAR_INPUT
		SourceDest 	: t_SourceDest;
		pNewPDO 	: ^t_PDOElement;
	END_VAR
	VAR_OUTPUT
		pRecyclePDO 	: ^t_PDOElement;
	END_VAR
  VAR
  	i : UDINT;
    pHelpInfo : ^t_PDOModuleInfo;
    pSearchInfo : ^t_PDOModuleInfo;
    ppHelpManaging : ^t_pManagingComponent;
    pSearchManaging : ^t_ManagingComponent;
  END_VAR

  // initialize with invalid
  pRecyclePDO := NIL;

  // if we have no pdoelements yet, quit
  if PDOElementNo = 0 then
    return;
  end_if;

  // we search for a PDO with the same source (then it contains the same data)
  pHelpInfo := #aPDOElements[0].SourceInfo;
  pSearchInfo := #pNewPDO^.SourceInfo;

  case SourceDest of
    SourceDest_IsSource:
      ppHelpManaging := #aPDOElements[0].pManagingSource;
      pSearchManaging := pNewPDO^.pManagingSource;
    SourceDest_IsDest:
      ppHelpManaging := #aPDOElements[0].pManagingDest;
      pSearchManaging := pNewPDO^.pManagingDest;
  else
    return;
  end_case;

  // check if we already have the path info of this source/destination
  for i := 0 to (PDOElementNo-1) do
    // if managing node, pathlength and path matches
    if (ppHelpManaging^ = pSearchManaging) & (pHelpInfo^.PathLen = pSearchInfo^.PathLen) & (To_StdLib.MemCmp(pHelpInfo^.pPath, pSearchInfo^.pPath, pHelpInfo^.PathLen) = 0) then
      // we found our PDO to recycle (PDO is already tranferred over this managing node
      pRecyclePDO := #aPDOElements[i];
      return;
    end_if;

    pHelpInfo       += sizeof(t_PDOElement);
    ppHelpManaging  += sizeof(t_PDOElement);
  end_for;

END_FUNCTION

FUNCTION SafetyManager::AddManagingInfo
	VAR_INPUT
		pPara 	: ^CmdStruct;
	END_VAR
  VAR
  	pHelpManaging : ^t_ManagingComponent;
  END_VAR

(*
  Parameter description:
  0..pointer to write PDOs in VARAN manager DPRAM
  1..pointer to read PDOs in VARAN manager DPRAM
  2..thispointer of calling class
  3..pointer to write PDOs in internal memory
  4..pointer to read PDOs in internal memory
  5..maximum available space for write PDOs in bytes
  6..maximum available space for read PDOs in bytes
*)

  pHelpManaging := pFirstManagingInterfaceComponent;
  while pHelpManaging do
    if pHelpManaging^.pThis = pPara^.aPara[2]$pVirtualBase then
      exit;
    end_if;

    pHelpManaging := pHelpManaging^.pNext;
  end_while;

  if pHelpManaging then
    pHelpManaging^.pPDOWriteSpaceDPRAM  := pPara^.aPara[0]$^USINT;
    pHelpManaging^.pPDOReadSpaceDPRAM   := pPara^.aPara[1]$^USINT;

    pHelpManaging^.pPDOWriteSpace       := pPara^.aPara[3]$^USINT;
    pHelpManaging^.pPDOReadSpace        := pPara^.aPara[4]$^USINT;

    pHelpManaging^.PDOWriteMemAvailable := pPara^.aPara[5]$UDINT;
    pHelpManaging^.PDOReadMemAvailable  := pPara^.aPara[6]$UDINT;

    pHelpManaging^.ud_HandlePDOWriteSpaceDPRAM  := pPara^.aPara[7]$UDINT;
    pHelpManaging^.ud_HandlePDOReadSpaceDPRAM   := pPara^.aPara[8]$UDINT;

  end_if;

END_FUNCTION

FUNCTION SafetyManager::CheckModuleUsage
	VAR_INPUT
		Length 	: UINT;
		pData 	: ^void;
		IsFSoEConfig 	: BOOL;
	END_VAR
	VAR_OUTPUT
		retcode 	: DINT;
	END_VAR
  VAR
    pDataHelp : ^void;
    i : UDINT;
    TmpPathLen : UINT;
    TempCfgNo : USINT;
    ModuleCfgInfo : t_ModuleCfgInfo;
    PdoCfgInfo : t_PdoCfgInfo;
    TempConnectionNo : UINT;
  END_VAR

(*
    Memory structure:
      4 Byte: SafetyNumber of CPU (is already there from initialisation in CSCP011_IM::InitSafeModule)
      1 Byte: Number of module configurations which are following
      for every module configuration (first is always the CPU itself)
        1 Byte: Info
        4 Byte: Interface Frame Source SafetyNumber (0 if it is no source for interface frames)
        4 Byte: Interface Frame CRC
        1 Byte: Number of destination inferface frame CRCs
        x Byte: Destination interface frame CRCs (number * sizeof(HDINT)
        2 Byte: Length of hardware path
        x Byte (depending on length in the 2 byte before): Hardwarepath
        2 Byte: Length of compressed hardware path
        x Byte (depending on length in the 2 byte before): Compressed Hardwarepath
        1 Byte: PDO out length for this module
      1 Byte: Number of pdo configurations which are following
      for every PDO configuration
        1 Byte: PDO length
        1 Byte: Interface frame info
        4 Byte: Interface CRC
        2 Byte: Length of source hardware path
        x Byte (depending on length in the 2 byte before): Hardwarepath of source
        2 Byte: Length of destination hardware path
        x Byte (depending on length in the 2 byte before): Hardwarepath of destination
      1 Byte: Number of slave configurations which are following
      for every slave configuration
        1 Byte: Info
        4 Byte: InterfaceCRC
        2 Byte: Length of hardware path
        x Byte (depending on length in the 2 byte before): Hardwarepath
        2 Byte: Length of compressed hardware path
        x Byte (depending on length in the 2 byte before): Compressed Hardwarepath

      if IsFSoEConfig = TRUE
      2 Byte: Number of connection infos which are following
      for every FSoE connection info
        2 Byte: ConnectionID
        1 Byte: ConnectionState
        1 Byte: Flags
        4 Byte: Master safety number
        2 Byte: Offset where to read from master
        2 Byte: Size of data to read from master (and write to slave)
        2 Byte: Offset where to write to master
        2 Byte: Size of data to write to master (and read from slave)
        2 Byte: SlaveAddress
        2 Byte: Length of slave hardware path
        x Byte (depending on length in the 2 byte before): Slave hardware path
        2 Byte: Length of compressed slave hardware path
        x Byte (depending on length in the 2 byte before): Compressed slave hardware path
        2 Byte: Offset where to read from slave
        2 Byte: Offset where to write to slave
*)

  // check if the configuration is valid (pData <> NIL) & (Length must be at least 4 byte for SafetyNbr + 1 byte module cfg number + 1 byte pdo cfg number + 1 byte slave cfc number)
  if pData & (Length >= 7)  then

    retcode := 0;

    pDataHelp := pData;

    // skip safety number of the safety cpu
    pDataHelp += sizeof(HDINT);

    // number of module configurations which follow now
    TempCfgNo := pDataHelp^$USINT;

    // skip number of module configurations
    pDataHelp += sizeof(USINT);

    // module configurations
    if TempCfgNo then
      for i := 0 to (TempCfgNo-1) do
        // info
        ModuleCfgInfo := pDataHelp^$t_ModuleCfgInfo;

        // skip info
        pDataHelp += sizeof(BSINT);

        // skip safety number of interface frame source
        pDataHelp += sizeof(HDINT);

        // skip interface CRC of interface frame
        pDataHelp += sizeof(HDINT);

        // interface frame destination CRCs
        if ModuleCfgInfo.IsInterfaceDest then
          // number of CRCs
          TmpPathLen := pDataHelp^$USINT;

          // skip number of CRCs
          pDataHelp += sizeof(USINT);

          // skip interface destination CRCs
          pDataHelp += TmpPathLen * sizeof(HDINT);
        end_if;

        // length of hardware path
        TmpPathLen := pDataHelp^$UINT;

        // skip length of hardware path
        pDataHelp += sizeof(UINT);

        SetModuleUsed(PathLen:=TmpPathLen, pPath:=pDataHelp$^USINT, IgnoreOptional:=FALSE, IsOptional:=ModuleCfgInfo.IsOptional, IsInterfaceDomain := FALSE);

        // skip hardware path
        pDataHelp += TmpPathLen;

        // length of compressed hardware path
        TmpPathLen := pDataHelp^$UINT; // save some time with this local variable

        // skip length of compressed hardware path
        pDataHelp += sizeof(UINT);

        // skip compressed hardware path
        pDataHelp += TmpPathLen;

        // skip pdo out length of this module
        pDataHelp += sizeof(USINT);
      end_for;
    end_if;

    // number of Pdo configurations which follow now
    TempCfgNo := pDataHelp^$USINT;

    // skip number of pdo configurations
    pDataHelp += sizeof(USINT);

    // Pdo configurations
    if TempCfgNo then
      for i := 0 to (TempCfgNo-1) do
        // skip pdo length
        pDataHelp += sizeof(USINT);

        // is it an interface pdo?
        PdoCfgInfo := pDataHelp^$t_PdoCfgInfo;

        // skip info
        pDataHelp += sizeof(BSINT);

        // skip interface CRC
        pDataHelp += sizeof(HDINT);

        // length of source hardware path
        TmpPathLen := pDataHelp^$UINT;

        // skip length of source hardware path
        pDataHelp += sizeof(UINT);

        SetModuleUsed(PathLen:=TmpPathLen, pPath:=pDataHelp$^USINT, IgnoreOptional:=FALSE, IsOptional:=PdoCfgInfo.IsOptional, IsInterfaceDomain := PdoCfgInfo.IsInterfacePDO);

        // skip source hardware path
        pDataHelp += TmpPathLen;

        // length of destination hardware path
        TmpPathLen := pDataHelp^$UINT;

        // skip length of destination hardware path
        pDataHelp += sizeof(UINT);

        // a destination module doesn't influence the optional property=> ignore the optional setting
        SetModuleUsed(PathLen:=TmpPathLen, pPath:=pDataHelp$^USINT, IgnoreOptional:=TRUE, IsOptional:=FALSE, IsInterfaceDomain := PdoCfgInfo.IsInterfacePDO);

        // skip destination hardware path
        pDataHelp += TmpPathLen;
      end_for;
    end_if;

    // number of slave configurations which follow now
    TempCfgNo := pDataHelp^$USINT;

    // skip number of slave configurations
    pDataHelp += sizeof(USINT);

    // slave configurations
    if TempCfgNo then
      for i := 0 to (TempCfgNo-1) do
        // skip info
        pDataHelp += sizeof(BSINT);

        // skip InterfaceCRC
        pDataHelp += sizeof(HDINT);

        // length of hardwarepath
        TmpPathLen := pDataHelp^$UINT; // save some time with this local variable

        // skip length of hardwarepath
        pDataHelp += sizeof(UINT);

        // skip hardwarepath
        pDataHelp += TmpPathLen;

        // length of compressed hardwarepath
        TmpPathLen := pDataHelp^$UINT; // save some time with this local variable

        // skip length of compressed hardwarepath
        pDataHelp += sizeof(UINT);

        // skip compressed hardwarepath
        pDataHelp += TmpPathLen;
      end_for;
    end_if;

    // check if it's a FSoE Config
    if IsFSoEConfig then
      // number of connection details which follow now
      TempConnectionNo := pDataHelp^$UINT;
      pDataHelp += sizeof(UINT);

      // if we got connections
      if TempConnectionNo then
        for i := 0 to (TempConnectionNo-1) do
          // connection ID
          pDataHelp += sizeof(UINT);

          // connection state
          pDataHelp += sizeof(USINT);

          // flags
          pDataHelp += sizeof(USINT);

          // master safety number
          pDataHelp += sizeof(HDINT);

          // offset where to read from master
          pDataHelp += sizeof(UINT);

          // size of data to read from master (and write to slave)
          pDataHelp += sizeof(UINT);

          // offset where to write to master
          pDataHelp += sizeof(UINT);

          // size of data to write to master (and read from slave)
          pDataHelp += sizeof(UINT);

          // slave address
          pDataHelp += sizeof(UINT);

          // length of uncompressed slave hardwarepath
          TmpPathLen := pDataHelp^$UINT; // save some time with this local variable
          pDataHelp += sizeof(UINT);

          // uncompressed slave hardwarepath
          pDataHelp += TmpPathLen;

          // length of compressed slave hardwarepath
          TmpPathLen := pDataHelp^$UINT; // save some time with this local variable
          pDataHelp += sizeof(UINT);

          // compressed slave hardwarepath
          pDataHelp += TmpPathLen;

          // offset where to read from master
          pDataHelp += sizeof(UINT);

          // offset where to write to master
          pDataHelp += sizeof(UINT);
        end_for;
      end_if;
    end_if;

    // check if the given size matches the memory structure
    if (pDataHelp$UDINT - pData$UDINT) <> Length then
      LogError("(SafetyManager::CheckModuleUsage) Invalid configuration data given (length doesn't match memory structure)");
      retcode := -3;
      return;
    end_if;
  else
    // invalid configuration
    LogError("(SafetyManager::CheckModuleUsage) Found invalid safety cpu configuration: Pointer or size wrong");
    retcode := -1;
  end_if;

END_FUNCTION

FUNCTION SafetyManager::SetModuleUsed
	VAR_INPUT
		PathLen 	: UINT;
		pPath 	: ^USINT;
		IgnoreOptional 	: BOOL;
		IsOptional 	: BOOL;
		IsInterfaceDomain 	: BOOL;
	END_VAR
  VAR
    pHelpManaging : ^t_ManagingComponent;
    pHelpSafety : ^t_SafetyComponent;
    TempPath : ARRAY [0..99] OF USINT;
  END_VAR

  // search for the hardware path

  // start with the safety components
  pHelpSafety := pFirstSafetyComponent;
  while pHelpSafety & pHelpSafety^.pPath do
    // we have 1 byte path length on the safety component but we got a 2 byte path length from the configuration
    // furthermore the pPath string could be over more domains and we have only our local path => check if length is bigger and if there is a domain escape right before the domain number
    if ((pPath^ = pHelpSafety^.pPath^) | ((pPath^ > pHelpSafety^.pPath^) & ((pPath + 1 + pPath^ - pHelpSafety^.pPath^)^ = HWT_ESCAPE_DOMAIN))) &
       (To_StdLib.MemCmp(pHelpSafety^.pPath + 1, pPath + 2 + pPath^ - pHelpSafety^.pPath^, pHelpSafety^.pPath^) = 0) then
      // only set IsOptional to false (has been initialized with true)
      if (IsOptional = FALSE) & (IgnoreOptional = FALSE) then
        pHelpSafety^.InfoBits.IsOptional := FALSE;
      end_if;
      return;
    end_if;

    pHelpSafety := pHelpSafety^.pNext;
  end_while;

  // if not found, continue with the managing interface components
  pHelpManaging := pFirstManagingInterfaceComponent;
  while pHelpManaging do
    if (To_StdLib.MemCmp(pHelpManaging^.pModulePath, pPath, PathLen) = 0) then
      // only set IsOptional to false (has been initialized with true)
      if (IsOptional = FALSE) & (IgnoreOptional = FALSE) then
        pHelpManaging^.InfoBits.IsOptional := FALSE;
      end_if;
      return;
    end_if;

    pHelpManaging := pHelpManaging^.pNext;
  end_while;

  _memcpy(ptr1:=#TempPath[0], ptr2:=pPath, cntr:=PathLen$USINT);

END_FUNCTION

FUNCTION SafetyManager::CreateTimeSyncList
  VAR
  	pHelp : ^t_TimeSyncElement;
  	pHelpSafety   : ^t_SafetyComponent;
  	pHelpManaging : ^t_ManagingComponent;
  END_VAR

  // first we stop time syncing (if active) to prevent crashing due tue a running time synchronisation
  pActTimeSyncElement := NIL;

  // if there is an old list, free it first
  if pFirstTimeSyncElement then
    // open the ring (set the next pointer of the last element to NIL)
    pFirstTimeSyncElement^.pPrev^.pNext := NIL;

    // remove the elements
    while pFirstTimeSyncElement do
      pHelp := pFirstTimeSyncElement;
      pFirstTimeSyncElement := pFirstTimeSyncElement^.pNext;

      To_StdLib.Free(mptr:=pHelp);
    end_while;
  end_if;

  pHelpSafety := pFirstSafetyComponent;
  while pHelpSafety do
    // if it's a module with not only inputs (then there's nothing to synchronize with) => trigger it for time synchronisation
    if (pHelpSafety^.InfoBits.OnlyInputs = FALSE) & (IsFSoEModule(pHelpSafety^.ModuleType) = FALSE) then
      AddTimeSyncElement(pManaging:=NIL, pSafety:=pHelpSafety, IsInterfaceDomain := FALSE);
    end_if;

    pHelpSafety := pHelpSafety^.pNext;
  end_while;

  // interface domains will not get our token, they got their own
  pHelpManaging := pFirstManagingInterfaceComponent;
  while pHelpManaging do
    AddTimeSyncElement(pManaging:=pHelpManaging, pSafety:=NIL, IsInterfaceDomain := TRUE);

    pHelpManaging := pHelpManaging^.pNext;
  end_while;

END_FUNCTION

FUNCTION SafetyManager::AddTimeSyncElement
	VAR_INPUT
		pManaging 	: ^t_ManagingComponent;
		pSafety 	: ^t_SafetyComponent;
		IsInterfaceDomain 	: BOOL;
	END_VAR
  VAR
    pLast : ^t_TimeSyncElement;
  	pHelp : ^t_TimeSyncElement;
  END_VAR

  // first we have to allocate some memory for the new element
  if pFirstTimeSyncElement = NIL then
    pFirstTimeSyncElement$pVoid := To_StdLib.Malloc(size:=sizeof(t_TimeSyncElement));
    pLast := pHelp := pFirstTimeSyncElement;
  else
    // check if we got this already
    pHelp := pFirstTimeSyncElement;
    repeat
      if pSafety & (pHelp^.pSafety = pSafety) then
        // already in list => leave
        return;
      end_if;

      if pManaging & (pHelp^.pManaging = pManaging) then
        // already in list => leave
        return;
      end_if;

      pHelp := pHelp^.pNext;
    until (pHelp = pFirstTimeSyncElement) end_repeat;

    pHelp$pVoid := To_StdLib.Malloc(size:=sizeof(t_TimeSyncElement));
    pLast := pFirstTimeSyncElement^.pPrev;
  end_if;

  if pHelp then
    // close the double linked ring with the new elements
    pFirstTimeSyncElement^.pPrev := pHelp;
    pHelp^.pNext := pFirstTimeSyncElement;

    pHelp^.pPrev := pLast;
    pLast^.pNext := pHelp;

    pHelp^.InfoBits := 0;
    pHelp^.InfoBits.IsInterfaceDomain := IsInterfaceDomain;

    pHelp^.pManaging := pManaging;
    pHelp^.pSafety   := pSafety;

    // managing modules
    if (pManaging <> NIL) then
      pHelp^.InfoBits.IsManagingModule := TRUE;
      pHelp^.pThis := pManaging^.pThis;

      // if it's the master connection
      if pManaging^.InfoBits.IsConnectionToMaster then
        // remember it
        pHelp^.InfoBits.IsConnectionToMaster := TRUE;

        // and make it the end of the list
        pFirstTimeSyncElement := pHelp^.pNext;

        // remember that we got a master connection
        pMasterTimeSyncElement := pHelp;

      elsif pMasterTimeSyncElement then
        // if we're not master and there is already a master time sync element in the list, we have to make it the last element
        pFirstTimeSyncElement := pMasterTimeSyncElement^.pNext;
      end_if;
    else
      // safety modules
      pHelp^.InfoBits.IsManagingModule := FALSE;
      pHelp^.pThis := pSafety^.pThis;

    // insert new safety modules at the beginning (managing modules at the end)
      pFirstTimeSyncElement := pHelp;
    end_if;

  else
    ClassState := -1;
    LogError("(SafetyManager::AddTimeSyncElement) Failed to allocate memory for a new Element");
  end_if;

END_FUNCTION

FUNCTION SafetyManager::CreateVirtualPDOs
  VAR
  	pHelpManaging   : ^t_ManagingComponent;
    pHelpConfig     : ^t_CfgListElem;
    pHelpPdo        : ^t_PdoListElem;
    TempPDO         : t_PdoCfg;
    pSearchConfig   : ^t_CfgListElem;
    pSearchPdo      : ^t_PdoListElem;
    b_UsedAsDest    : BOOL;
  END_VAR

  pHelpConfig := pConfigs;
  while pHelpConfig do
    pHelpPdo := pHelpConfig^.pFirstPdoCfg;
    while pHelpPdo do
      // check if it's a broadcast
      if (pHelpPdo^.PdoInfo.Info.IFBroadCast) & (pHelpPdo^.PdoInfo.Info.VirtualPDOsCreated = FALSE) then
        // found one => create virtual PDOs from it (add them to the same configuration)

        // prepare new virtual PDO
        TempPDO := pHelpPdo^.PdoInfo;

        TempPDO.Info.IFBroadCast := FALSE;
        TempPDO.Info.VirtualPDO := TRUE;

        // add a new PDO for every interface managing module
        pHelpManaging := pFirstManagingInterfaceComponent;
        while pHelpManaging do
          // change destination path to the actual module
          TempPDO.DestPathLen := pHelpManaging^.pModulePath^ + 2;
          TempPDO.pDestPath := pHelpManaging^.pModulePath;

          if AddVirtualPDOToCfg(pCfg:=pHelpConfig, pNewPDO:=#TempPDO) then
            LogError(e_msg:="(SafetyManager::CreateVirtualPDOs) Failed to allocate memory for a new virtual PDO");
          end_if;

          pHelpManaging := pHelpManaging^.pNext;
        end_while;

        // search in all configs (if there are other) for a pdo with this interface CRC as source
        pSearchConfig := pConfigs;
        while pSearchConfig do
          pSearchPdo := pSearchConfig^.pFirstPdoCfg;
          while pSearchPdo do
            // we must not manipulate our help pdo
            if pSearchPdo <> pHelpPdo then
              b_UsedAsDest := FALSE;

              // check if the path is already used as destination
              if (pSearchPdo^.PdoInfo.DestPathLen = pHelpPdo^.PdoInfo.SourcePathLen) &
                 (To_StdLib.MemCmp(pSearchPdo^.PdoInfo.pDestPath, pHelpPdo^.PdoInfo.pSourcePath, pHelpPdo^.PdoInfo.SourcePathLen) = 0) then
                b_UsedAsDest := TRUE;
              end_if;

              // check if the interface CRC appears in any PDO (only if the path isn't already used as destination path)
              if (pSearchPdo^.PdoInfo.InterfaceCRC = pHelpPdo^.PdoInfo.InterfaceCRC) & (b_UsedAsDest = FALSE) then
                // now take the source path of the broadcast PDO and use it as source path for this PDO
                To_StdLib.Free(mptr:=pSearchPdo^.PdoInfo.pSourcePath);

                pSearchPdo^.PdoInfo.pSourcePath$pVoid := To_StdLib.Malloc(size:=pHelpPdo^.PdoInfo.SourcePathLen);

                // save source hardwarepath
                if pSearchPdo^.PdoInfo.pSourcePath then
                  _memcpy(ptr1:=pSearchPdo^.PdoInfo.pSourcePath, ptr2:=pHelpPdo^.PdoInfo.pSourcePath, cntr:=pHelpPdo^.PdoInfo.SourcePathLen);
                  pSearchPdo^.PdoInfo.SourcePathLen := pHelpPdo^.PdoInfo.SourcePathLen;

                  // source and destination of this PDO are both local safe cpu modules which communicate with each other via interface frames => store them in extra list for routing SDOs and TDOs
                  AddToLocalIFs(#pSearchPdo^.PdoInfo);
                else
                  LogError(e_msg:="(SafetyManager::CreateVirtualPDOs) Failed to allocate memory for a source path");
                  pSearchPdo^.PdoInfo.SourcePathLen := 0;
                  ClassState := -1;
                end_if;
              end_if;
            end_if;

            pSearchPdo := pSearchPdo^.pNext;
          end_while;

          pSearchConfig := pSearchConfig^.pNext;
        end_while;
        pHelpPdo^.PdoInfo.Info.VirtualPDOsCreated := TRUE;
      end_if;

      pHelpPdo := pHelpPdo^.pNext;
    end_while;

    pHelpConfig := pHelpConfig^.pNext;
  end_while;

END_FUNCTION

FUNCTION SafetyManager::AddVirtualPDOToCfg
	VAR_INPUT
		pCfg 	: ^t_CfgListElem;
		pNewPDO 	: ^t_PdoCfg;
	END_VAR
	VAR_OUTPUT
		retcode 	: DINT;
	END_VAR
  VAR
    pHelpPdo        : ^t_PdoListElem;
    TempLen         : UINT;
  END_VAR

  retcode := 0;

  if pCfg^.pFirstPdoCfg = NIL then
    // first PDO in this cfg (should not be possible, because the template for this PDO is also in the same config)
    pCfg^.pFirstPdoCfg$pVoid := To_StdLib.Malloc(size:=sizeof(t_PdoListElem));
    pHelpPdo := pCfg^.pFirstPdoCfg;
  else
    // search a place for the new PDO
    pHelpPdo := pCfg^.pFirstPdoCfg;
    while pHelpPdo^.pNext do

      pHelpPdo := pHelpPdo^.pNext;
    end_while;

    pHelpPdo^.pNext$pvoid := To_StdLib.Malloc(size:=sizeof(t_PdoListElem));
    pHelpPdo := pHelpPdo^.pNext;
  end_if;

  if pHelpPdo then
    // init the values
    pHelpPdo^.PdoInfo.PdoLen        := pNewPDO^.PdoLen;
    pHelpPdo^.PdoInfo.Info          := pNewPDO^.Info;
    pHelpPdo^.PdoInfo.InterfaceCRC  := pNewPDO^.InterfaceCRC;

    // length of source hardwarepath
    TempLen := pNewPDO^.SourcePathLen; // save some time with this local variable
    pHelpPdo^.PdoInfo.SourcePathLen := TempLen;

    // allocate memory for the source module path
    pHelpPdo^.PdoInfo.pSourcePath$pVoid := To_StdLib.Malloc(size:=TempLen);
    if pHelpPdo^.PdoInfo.pSourcePath = NIL then
      ClassState := -1;
      retcode := -2;
      return;
    end_if;

    // save source hardwarepath
    _memcpy(ptr1:=pHelpPdo^.PdoInfo.pSourcePath, ptr2:=pNewPDO^.pSourcePath, cntr:=TempLen);

    // length of destination hardwarepath
    TempLen := pNewPDO^.DestPathLen; // save some time with this local variable
    pHelpPdo^.PdoInfo.DestPathLen := TempLen;

    // allocate memory for the destination module path
    pHelpPdo^.PdoInfo.pDestPath$pVoid := To_StdLib.Malloc(size:=TempLen);
    if pHelpPdo^.PdoInfo.pDestPath = NIL then
      ClassState := -1;
      retcode := -2;
      return;
    end_if;

    // save destination hardwarepath
    _memcpy(ptr1:=pHelpPdo^.PdoInfo.pDestPath, ptr2:=pNewPDO^.pDestPath, cntr:=TempLen);

    // now we give it an ID and increase the number for the next pdo
    pHelpPdo^.PdoInfo.PDO_ID := ActPDO_ID;
    ActPDO_ID += 1;

    pHelpPdo^.pNext                  := NIL;
  else
    ClassState := -1;
    retcode := -2;
    return;
  end_if;

END_FUNCTION

FUNCTION SafetyManager::AddToLocalIFs
	VAR_INPUT
		pHelpPDO 	: ^t_PdoCfg;
	END_VAR
  VAR
  	AddSource : BOOL;
    i : USINT;
    pHelpSafety : ^t_SafetyComponent;
  END_VAR

  // check if there is still room for new modules
  if LocalIFNo < MAX_INTERNAL_IF_MODULES then

    AddSource := TRUE;

    // if there is a list, check if any of our modules are already in the list
    if LocalIFNo then
      for i := 0 to (LocalIFNo-1) do
        // check if crc matches
        if (aLocalIFs[i].InterfaceCRC = pHelpPDO^.InterfaceCRC) then
          AddSource := FALSE;
          exit;
        end_if;
      end_for;
    end_if;

    // now we know how many we have to add to the list. if there are modules to add and there is enough space for all of them => do it
    if AddSource then
      // search it in the local modules
      pHelpSafety := pFirstSafetyComponent;
      while pHelpSafety do
        // if the path matches, add the module to the list

        // source module
        if (pHelpSafety^.PathLen = (pHelpPDO^.SourcePathLen - 1)) &
        // we compare the last x byte (where x is the length of the local path including the domain) because we got different length info sizes (1 byte vs. 2 byte)
           (To_StdLib.MemCmp(pHelpSafety^.pPath + 1, pHelpPDO^.pSourcePath + 2 + pHelpPDO^.pSourcePath^ - pHelpSafety^.pPath^, pHelpSafety^.pPath^) = 0) then
          aLocalIFs[LocalIFNo].InterfaceCRC  := pHelpPDO^.InterfaceCRC;
          aLocalIFs[LocalIFNo].pSafetyModule := pHelpSafety;
          LocalIFNo += 1;
          exit;
        end_if;

        pHelpSafety := pHelpSafety^.pNext;
      end_while;
    end_if;
  end_if;

END_FUNCTION

FUNCTION SafetyManager::IFInfoNotArrivedYet
	VAR_INPUT
		pThis 	: pVirtualBase;
	END_VAR
	VAR_OUTPUT
		InfoNotAvailable 	: BOOL;
	END_VAR
  VAR
  	pHelpManaging : ^t_ManagingComponent;
  END_VAR

	InfoNotAvailable := FALSE;

  pHelpManaging := pFirstManagingInterfaceComponent;
  while pHelpManaging do
    if pHelpManaging^.pThis = pThis then
      if pHelpManaging^.InfoBits.GotIFInfo = FALSE then
        InfoNotAvailable := TRUE;
      end_if;
      return;
    end_if;

    pHelpManaging := pHelpManaging^.pNext;
  end_while;

END_FUNCTION

#pragma warning(disable:74)
FUNCTION SafetyManager::StartTimeMeasurement
	VAR_INPUT
		usMode (EAX) 	: DINT;
	END_VAR
#ifdef VM_CLASS_TIME_MEASUREMENT
  VAR
  	tmpTime : ^t_TimeMeasurementVaran;
  END_VAR

  case usMode of

    //-----------------------------------------------------------

    VARANTIME_RT:
      tmpTime := #s_TimeRt;

    //-----------------------------------------------------------

    VARANTIME_RTPOSTSCAN:
      tmpTime := #s_TimeRtPostScan;

    //-----------------------------------------------------------

    VARANTIME_CY:
      tmpTime := #s_TimeCy;

    //-----------------------------------------------------------

  end_case;

  if ( tmpTime^.us_Activate ) then
//    Save_Flg();
//    CLI();
    tmpTime^.ud_Timemark := OS_READMICROSEC();
  end_if;

#endif

END_FUNCTION

FUNCTION SafetyManager::StopTimeMeasurement
	VAR_INPUT
		usMode (EAX) 	: DINT;
	END_VAR
#ifdef VM_CLASS_TIME_MEASUREMENT
  VAR
  	tmpTime : ^t_TimeMeasurementVaran;
  END_VAR

  case usMode of

    //-----------------------------------------------------------

    VARANTIME_RT:
      tmpTime := #s_TimeRt;

    //-----------------------------------------------------------

    VARANTIME_RTPOSTSCAN:
      tmpTime := #s_TimeRtPostScan;

    //-----------------------------------------------------------

    VARANTIME_CY:
      tmpTime := #s_TimeCy;

    //-----------------------------------------------------------

  end_case;

	if ( tmpTime^.us_Activate ) then

		//get actual time
		tmpTime^.ud_ActualTime := OS_READMICROSEC();
    tmpTime^.ud_ActualTime -= tmpTime^.ud_Timemark;

		//look for maximum time
		if ( tmpTime^.ud_ActualTime > tmpTime^.ud_MaximalTime ) then
			tmpTime^.ud_MaximalTime := tmpTime^.ud_ActualTime;
		end_if;

		//look for minimum time
		if ( tmpTime^.ud_ActualTime < tmpTime^.ud_MinimalTime ) then
			tmpTime^.ud_MinimalTime := tmpTime^.ud_ActualTime;
		end_if;

		//look for average time (100000 cycles)
		if ( tmpTime^.ud_AverageCounter = 100000 ) then

			tmpTime^.ud_AverageTime 	:= tmpTime^.ud_AverageSum / tmpTime^.ud_AverageCounter;
			tmpTime^.ud_AverageSum 	:= 0;
			tmpTime^.ud_AverageCounter := 0;

		else
			tmpTime^.ud_AverageSum += ( tmpTime^.ud_ActualTime / 100 );
			tmpTime^.ud_AverageCounter += 1;
		end_if;

//		STI();
//    Restore_Flg();
	end_if;

#endif

END_FUNCTION // Varan_Base::StopTimeMeasurement
#pragma warning(default:74)

FUNCTION SafetyManager::AnyIFDomainSynchron
	VAR_OUTPUT
		AnythingSynchron 	: BOOL;
	END_VAR
  VAR
    pHelpManaging   : ^t_ManagingComponent;
  END_VAR

  AnythingSynchron := FALSE;

  pHelpManaging := pFirstManagingInterfaceComponent;
  while pHelpManaging do
    if pHelpManaging^.InfoBits.IsSynchron then
      AnythingSynchron := TRUE;
      return;
    end_if;

    pHelpManaging := pHelpManaging^.pNext;
  end_while;

END_FUNCTION

FUNCTION SafetyManager::LocalIFsAvailable
	VAR_OUTPUT
		retcode 	: BOOL;
	END_VAR
  VAR
    pHelpCfg : ^t_CfgListElem;
    pHelpPdo : ^t_PdoListElem;
    pHelpModule : ^t_ModuleListElem;
  END_VAR

  retcode := FALSE;

  // add all local configs to our structure
  SendLocalCfgsToMaster();

  // check the local configs for interface frames
  pHelpCfg := pConfigs;
  while pHelpCfg do
    pHelpPdo := pHelpCfg^.pFirstPdoCfg;
    while pHelpPdo do
      if pHelpPdo^.PdoInfo.Info.IsInterfacePDO | pHelpPdo^.PdoInfo.Info.IFBroadCast then
        retcode := TRUE;
        return;
      end_if;

      pHelpPdo := pHelpPdo^.pNext;
    end_while;

    pHelpModule := pHelpCfg^.pFirstModuleCfg;
    while pHelpModule do
      if pHelpModule^.ModuleInfo.Info.IsInterfaceSource | pHelpModule^.ModuleInfo.Info.IsInterfaceDest then
        retcode := TRUE;
        return;
      end_if;

      pHelpModule := pHelpModule^.pNext;
    end_while;

    pHelpCfg := pHelpCfg^.pNext;
  end_while;

END_FUNCTION

FUNCTION SafetyManager::IsCPUModule
  VAR_INPUT
    ModuleType : t_e_ModuleType;
  END_VAR
  VAR_OUTPUT
  	retcode : BOOL;
  END_VAR

  case ModuleType of
    _CSCP01x,
    _SCP010,
    _SCP011,
    _SCP111,
    _SDD1300,
    _SDD1400,
    _SDD1500,
    _SDD1600:
      retcode := TRUE;
  else
    retcode := FALSE;
  end_case;

END_FUNCTION

FUNCTION SafetyManager::IsFSoEModule
	VAR_INPUT
		ModuleType 	: t_e_ModuleType;
	END_VAR
	VAR_OUTPUT
		retcode 	: BOOL;
	END_VAR

  case ModuleType of
    _SCP111,
    _SDD1300,
    _SDD1400,
    _SDD1500,
    _SDD1600:
      retcode := TRUE;
  else
    retcode := FALSE;
  end_case;

END_FUNCTION

FUNCTION SafetyManager::CreateFSoEPDOs
  VAR
  	pHelpConfigManager      : ^t_CfgListElem;
    pHelpConnectionManager  : ^t_FSoEConnectionDetails;
  	pHelpConfigSlave        : ^t_CfgListElem;
    pHelpConnectionSlave    : ^t_FSoEConnectionDetails;
    SlavesFoundNo           : INT;
    pLastFoundSlave         : ^t_FSoEConnectionDetails;
    pLastFoundSlaveCfg      : ^t_CfgListElem;
    SortConnectionList      : BOOL;
    ConnectionsAvailable    : UINT;
    pConnectionPointerList  : pVoid;
    ActIndex                : UINT;
  END_VAR

//*****************************************************************************
//** SEARCH FOR MASTER / SLAVE PAIRS VIA SLAVE ADDRESS                       **
//*****************************************************************************

  SortConnectionList    := FALSE;
  ConnectionsAvailable  := 0;

  // check all configs for manager connections (those contain the info about the slaves)
  pHelpConfigManager := pConfigs;
  while pHelpConfigManager do

    pHelpConnectionManager := pHelpConfigManager^.pFirstFSoEConnection;
    while pHelpConnectionManager do

      ConnectionsAvailable += 1;

      // if we got a master connection => search for a match of the slaveaddress in the slave configurations
      if pHelpConnectionManager^.Flags.IsMaster then
        SlavesFoundNo := 0;

        pHelpConfigSlave := pConfigs;
        while pHelpConfigSlave do

          pHelpConnectionSlave := pHelpConfigSlave^.pFirstFSoEConnection;
          while pHelpConnectionSlave do
            if pHelpConnectionSlave^.Flags.IsMaster = FALSE then
              if pHelpConnectionManager^.SlaveAddress = pHelpConnectionSlave^.SlaveAddress then
                // check if it's an internal interface frame
                if pHelpConnectionManager^.Flags.IsInterfaceConnection & pHelpConnectionSlave^.Flags.IsInterfaceConnection then
                  // check if the connection is still available
                  if pHelpConnectionSlave^.InternalConnectionState = FCS_RESET then
                    pLastFoundSlave     := pHelpConnectionSlave;
                    pLastFoundSlaveCfg  := pHelpConfigSlave;

                    // mark as internal interface frame
                    SlavesFoundNo := -1;

                    // exit both loops
                    pHelpConfigSlave := NIL;
                    exit;
                  end_if;
                else
                  SlavesFoundNo       += 1;
                  pLastFoundSlave     := pHelpConnectionSlave;
                  pLastFoundSlaveCfg  := pHelpConfigSlave;
                end_if;
              end_if;
            end_if;

            pHelpConnectionSlave := pHelpConnectionSlave^.pNext;
          end_while;

          if pHelpConfigSlave then
            pHelpConfigSlave := pHelpConfigSlave^.pNext;
          end_if;
        end_while;

        if SlavesFoundNo = 1 then
          // perfect, since the slave address is meant to be unique
          ShareConnectionInfos(pHelpConnectionManager, pHelpConfigManager, pLastFoundSlave, pLastFoundSlaveCfg);

        elsif SlavesFoundNo = 0 then
          // we have to search for the address in other systems which could be connected via interfaceframe
          if pFirstManagingInterfaceComponent = NIL then
            if pHelpConnectionManager^.SlaveAddress <> 0 then
              LogValue(pString:="(SafetyManager::CreateFSoEPDOs) Could not find Slave for Master connection with SlaveAddress 0x{0}", Value:=pHelpConnectionManager^.SlaveAddress);
            end_if;
          else
            SortConnectionList := TRUE;
          end_if;
        elsif SlavesFoundNo = -1 then
          // internal interface frame => add it to the list for SDO routing
          AddInternalIFFSoE(pHelpConnectionManager, pHelpConfigManager, pLastFoundSlave, pLastFoundSlaveCfg);
        else
          LogValue(pString:="(SafetyManager::CreateFSoEPDOs) Found more than 1 Slave for Master connection with SlaveAddress 0x{0}! Slave Address must be unique!", Value:=pHelpConnectionManager^.SlaveAddress);
        end_if;
      else
        if pHelpConnectionManager^.Flags.IsInterfaceConnection then
          if pFirstManagingInterfaceComponent then
            SortConnectionList := TRUE;
          end_if;

          // check if we can get an interface crc from the config
          if pHelpConfigManager^.pFirstModuleCfg & (pHelpConfigManager^.pFirstModuleCfg^.ModuleInfo.SafetyNbr = pHelpConnectionManager^.OwnerSafetyNbr) then
            // store the interface CRC (to send it to the other domain later)
            if pHelpConnectionManager^.pSlavePathComp = NIL then
              pHelpConnectionManager^.pSlavePathComp$pVoid := To_StdLib.Malloc(size:=8);

              if pHelpConnectionManager^.pSlavePathComp then
                // generate a compressed path (IF CRC)
                _memset(dest:=pHelpConnectionManager^.pSlavePathComp, usByte:=16#FF, cntr:=8);
                pHelpConnectionManager^.pSlavePathComp^$USINT := 3;
                _memcpy(ptr1:=pHelpConnectionManager^.pSlavePathComp + 1, ptr2:=#pHelpConfigManager^.pFirstModuleCfg^.ModuleInfo.InterfaceCRC, cntr:=sizeof(HDINT));
                pHelpConnectionManager^.SlavePathCompLen := 8;
              else
                LogError(e_msg:="(SafetyManager::CreateFSoEPDOs) Failed to allocate memory for an interface CRC!");
              end_if;
            end_if;
          end_if;
        end_if;
      end_if;

      pHelpConnectionManager := pHelpConnectionManager^.pNext;
    end_while;

    pHelpConfigManager := pHelpConfigManager^.pNext;
  end_while;

  // check if we got all slave addresses of local configs
  CheckLocalSlaveAddresses();

  // reset pointer
  pSortedConnections := NIL;

  // there are interface connections => sort the list by slave address to ensure correct order in memory
  if SortConnectionList | (ConnectionsAvailable & (b_AllLocalSlaveAddressesValid = FALSE)) then
    // first we need a pointer list of connection (not linked) with 4 byte entries
    pConnectionPointerList := To_StdLib.Malloc(size:=ConnectionsAvailable * sizeof(pVoid));

    if pConnectionPointerList = NIL then
      LogError(e_msg:="(SafetyManager::CreateFSoEPDOs) Failed to allocate memory for sorting the FSoE connections!");
      return;
    end_if;

    // store the pointers of all connections into the array
    ActIndex := 0;
    pHelpConfigManager := pConfigs;
    while pHelpConfigManager do

      pHelpConnectionManager := pHelpConfigManager^.pFirstFSoEConnection;
      while pHelpConnectionManager do
        (pConnectionPointerList + ActIndex * sizeof(pVoid))^$^t_FSoEConnectionDetails := pHelpConnectionManager;

        ActIndex                += 1;
        pHelpConnectionManager  := pHelpConnectionManager^.pNext;
      end_while;

      pHelpConfigManager := pHelpConfigManager^.pNext;
    end_while;

    // now that we got our linear memory to sort => do it
    MySort(src:=pConnectionPointerList$^USINT, no:=ActIndex, itemsize:=sizeof(pVoid), sortfunct:=#ConnectionSort());

    // create the new sorted linked list
    pSortedConnections := pConnectionPointerList^$^t_FSoEConnectionDetails;
    pHelpConnectionManager := pSortedConnections;

    // we already have the first connection at the pSortedConnections;
    for ActIndex := 1 to ConnectionsAvailable-1 do
      pHelpConnectionManager^.pNextSorted := (pConnectionPointerList + ActIndex * sizeof(pVoid))^$^t_FSoEConnectionDetails;
      pHelpConnectionManager := pHelpConnectionManager^.pNextSorted;
    end_for;

    To_StdLib.Free(mptr:=pConnectionPointerList);
    // now we can access the connection in order of the slave address via pSortedConnections
  end_if;

END_FUNCTION

FUNCTION SafetyManager::ShareConnectionInfos
	VAR_INPUT
		pMasterConnection 	: ^t_FSoEConnectionDetails;
		pMasterConfig 	: ^t_CfgListElem;
		pSlaveConnection 	: ^t_FSoEConnectionDetails;
		pSlaveConfig 	: ^t_CfgListElem;
	END_VAR
  VAR
  	pHelpSafety   : ^t_SafetyComponent;
    pMasterSafety : ^t_SafetyComponent;
    pSlaveSafety  : ^t_SafetyComponent;
		MyPara 	      : CmdStruct;
		MyResult	    : results;
    pPDOReadData  : pVoid;
    i             : UDINT;
    IsInList      : BOOL;
  END_VAR

//*****************************************************************************
//** TELL THE MODULES WHAT DATA TO COPY IN REALTIME                          **
//*****************************************************************************

  pMasterSafety := NIL;
  pSlaveSafety  := NIL;

  pHelpSafety := pFirstSafetyComponent;
  while pHelpSafety do

    if pHelpSafety^.SafetyNbr & (pHelpSafety^.SafetyNbr = pMasterConfig^.SafetyNbr) then
      pMasterSafety := pHelpSafety;
      exit;
    end_if;

    pHelpSafety := pHelpSafety^.pNext;
  end_while;

  pHelpSafety := pFirstSafetyComponent;
  while pHelpSafety do

    if pHelpSafety^.SafetyNbr & (pHelpSafety^.SafetyNbr = pSlaveConfig^.SafetyNbr) then
      pSlaveSafety := pHelpSafety;
      exit;
    end_if;

    pHelpSafety := pHelpSafety^.pNext;
  end_while;

  // if we found the safety modules who are keeping the configs => tell them what to copy
  if pMasterSafety & pSlaveSafety then
    // check for matching hardware paths
    if (pMasterConnection^.pSlavePath^ <> pSlaveSafety^.pPath^) |
       (To_StdLib.MemCmp(pSlaveSafety^.pPath + 1, pMasterConnection^.pSlavePath + 2, pSlaveSafety^.pPath^) <> 0) then
      LogError(e_msg:="(SafetyManager::ShareConnectionInfos) Error! The hardware path of the master connection doesn't match the hw path");
      LogValue(pString:=" of the slave module with the corresponding slave address (Slave Address 0x{0} and ConnectionID 0x{1})!", Value:=pMasterConnection^.SlaveAddress, Value2:=pMasterConnection^.ConnectionID);
      return;
    end_if;

    // check for equal sizes
    if (pMasterConnection^.MasterReadSize <> pSlaveConnection^.MasterReadSize) |
       (pMasterConnection^.MasterWriteSize <> pSlaveConnection^.MasterWriteSize) then
      LogError(e_msg:="(SafetyManager::ShareConnectionInfos) Error! The sizes of master and slave connection");
      LogValue(pString:="do not match for Slave Address 0x{0} and ConnectionID 0x{1}!", Value:=pMasterConnection^.SlaveAddress, Value2:=pMasterConnection^.ConnectionID);
      return;
    end_if;

    // we start with the safe outputs: get the data pointer from the master and give it to the slave
    MyPara.uiCmd    := CMD_SM_ADD_OUTPUT_PDO;
    MyResult.uiLng  := 0;
    pMasterSafety^.pThis^.NewInst(#MyPara, #MyResult);

    if MyResult.uiLng <> 4 then
      LogError(e_msg:="(SafetyManager::ShareConnectionInfos) Invalid return value when asking the master safety module for it's pointer to the PDO read data!");
      return;
    end_if;

    pPDOReadData := MyResult.aData[0]$pVoid;

#ifdef HWK_SHOW_PRAGMA_MESSAGES
#pragma message("RamAnd 20.11.2014 16:41 \ testweise mapping loggen")
    LogValue(pString:="(SafetyManager::ShareConnectionInfos) ConnectionID: {0}, SlaveAddress: {1}", Value:=pMasterConnection^.ConnectionID, Value2:=pMasterConnection^.SlaveAddress);
    LogValue(pString:="(SafetyManager::ShareConnectionInfos) MasterSafetyNbr: {0}, SlaveSafetyNbr: {1}", Value:=pMasterConnection^.OwnerSafetyNbr, Value2:=pSlaveConnection^.OwnerSafetyNbr);
    LogValue(pString:="(SafetyManager::ShareConnectionInfos) MasterReadOffset: {0}, MasterReadSize: {1}, SlaveWriteOffset: {2}", Value:=pMasterConnection^.MasterReadOffset, Value2:=pMasterConnection^.MasterReadSize, Value3 := pSlaveConnection^.SlaveWriteOffset);
#endif

    // check if it's in the list
    IsInList := FALSE;
    if FSoEInputPDONo then
      for i := 0 to FSoEInputPDONo do
        if ((aFSoEInputPDOs[i].pSafety = pSlaveSafety)  & (aFSoEInputPDOs[i].pMem = pPDOReadData$DINT + pMasterConnection^.MasterReadOffset)) then
          aFSoEInputPDOs[FSoEInputPDONo].pSafety    := pMasterSafety;
          aFSoEInputPDOs[FSoEInputPDONo].pMem       := MyPara.aPara[0];
          IsInList := TRUE;
        end_if;
      end_for;
    end_if;
